                   IF NOT #found THEN
                       #VarErr := 1;                       // no feasible transfer
                   ELSIF #CurLen >= 96 THEN
                       #VarErr := 2;                       // plan longer than 96 transfers
                   ELSE
                       // ---------- apply the best (s, d) ----------
                       #si := #bS;
                       #sCol := #SrcX[#si];
                       #sRow := #SrcY[#si];
                       #sBay := #SrcB[#si];
                       #dBay := #bDb;
                       #dCol := #FreeX[#dBay, #bK];
                       #dRow := #FreeY[#dBay, #bK];
                       #eT := "Crane_MoveCost"(X0 := #cx, Y0 := #cy, B0 := #cb, X1 := #sCol, Y1 := #sRow, B1 := #sBay,
                                               MMode := #cMMode, M => #eMan);
                       #lT := "Crane_MoveCost"(X0 := #sCol, Y0 := #sRow, B0 := #sBay, X1 := #dCol, Y1 := #dRow, B1 := #dBay,
                                               MMode := #cMMode, M => #lMan);
                       #g[#dBay, #dCol, #dRow] := #g[#sBay, #sCol, #sRow];
                       #g[#sBay, #sCol, #sRow] := 0;
                       #TotT := #TotT + #eT + 200 + #lT + 200;
                       #TotM := #TotM + INT_TO_DINT(#eMan) + 1 + INT_TO_DINT(#lMan) + 1;
                       #CurLen := #CurLen + 1;
                       #CurPlan[#CurLen].Kind := #SrcKind[#si];
                       #CurPlan[#CurLen].Id := #SrcId[#si];
                       #CurPlan[#CurLen].ListIdx := #SrcIdx[#si];
                       #CurPlan[#CurLen].SrcX := INT_TO_SINT(#sCol);
                       #CurPlan[#CurLen].SrcY := INT_TO_SINT(#sRow);
                       #CurPlan[#CurLen].SrcBay := INT_TO_USINT(#sBay);
                       #CurPlan[#CurLen].DstX := INT_TO_SINT(#dCol);
                       #CurPlan[#CurLen].DstY := INT_TO_SINT(#dRow);
                       #CurPlan[#CurLen].DstBay := INT_TO_USINT(#dBay);
                       #CurPlan[#CurLen].CumT_ds := #TotT;
                       #CurPlan[#CurLen].CumM := #TotM;
                       #CurSrc[#CurLen] := #si;
                       #cx := #dCol;
                       #cy := #dRow;
                       #cb := #dBay;
                       #cG := #FreeG[#dBay, #bK];
                       #Pend[#si] := FALSE;
                       #nPend := #nPend - 1;
                   END_IF;
               END_IF;

               IF #PubPending THEN
                   // ---------- job finished: publish (World is written only here) ----------
                   #PubPending := FALSE;
                   IF #HaveBest THEN
                       FOR #i := 1 TO 96 DO
                           IF #i <= #BestLen THEN
                               "World".Plan[#i] := #BestPlan[#i];
                           ELSE
                               "World".Plan[#i] := #ZeroTr;
                           END_IF;
                       END_FOR;
                       "World".PlanLen := #BestLen;
                       "World".PlanVariant := #BestV;
                       "World".PredT_ds := #BestT;
                       "World".PredM := #BestM;
                       "World".LbT_ds := #sBaseT + #LbT;
                       "World".LbM := #sBaseM + #LbM;
                       "World".ImpEvals := #ImpEvals;
                       "World".ImpAccepts := #ImpAcc;
                       "World".SlotAccepts := #SlAcc;
                       "World".OrderFeasible := #OrderOk;
                       IF #sN > 0 THEN
                           "World".PredJ := 0.5 * (DINT_TO_REAL(#BestT) / 10.0) / (76.0 * INT_TO_REAL(#sN))
                                          + 0.5 * DINT_TO_REAL(#BestM) / (4.0 * INT_TO_REAL(#sN));
                           "World".PredJ0 := 0.5 * (DINT_TO_REAL(#GrT) / 10.0) / (76.0 * INT_TO_REAL(#sN))
                                           + 0.5 * DINT_TO_REAL(#GrM) / (4.0 * INT_TO_REAL(#sN));
                           "World".LbJ := 0.5 * (DINT_TO_REAL(#sBaseT + #LbT) / 10.0) / (76.0 * INT_TO_REAL(#sN))
                                        + 0.5 * DINT_TO_REAL(#sBaseM + #LbM) / (4.0 * INT_TO_REAL(#sN));
                       ELSE
                           "World".PredJ := 0.0;
                           "World".PredJ0 := 0.0;
                           "World".LbJ := 0.0;
                       END_IF;
                       "World".PlanValid := TRUE;
                       #Done := TRUE;
                       #ErrCode := 0;
                   ELSE
                       "World".PlanValid := FALSE;
                       "World".PlanLen := 0;
                       "World".PlanVariant := 0;
                       "World".SlotAccepts := 0;
                       "World".OrderFeasible := #OrderOk;
                       #Error := TRUE;
                       #ErrCode := #Err1;
                   END_IF;
                   #JobBusy := FALSE;
               END_IF;
           END_WHILE;
           #DiagCallMs := RUNTIME(MEM := #RtMem) * 1000.0;
           #DiagJobMs := #DiagJobMs + #DiagCallMs;
           IF #DiagCallMs > #DiagMaxCallMs THEN
               #DiagMaxCallMs := #DiagCallMs;
           END_IF;
       END_IF;
   END_REGION

   #Busy := #JobBusy;
END_FUNCTION_BLOCK

FUNCTION "CheckCmd" : Int   // FC10, SCL
TITLE = Pre-check of a crane command before OB30 issues it to FB1
{ S7_Optimized_Access := 'TRUE' }
VERSION : 0.1
// Returns 0 = OK, otherwise the alarm bit number (CONTRACT 1.4 / 3.3):
//     100 ship imbalance (alarm bit 0)      1 pick location empty
//       2 drop location occupied            9 invalid command / position
//      11 crane already carrying (lift, or MANUAL reset with a load)   12 crane is empty (put down)
//   The first failing rule decides the result.
//   Lift/put act on the CURRENT crane position (CraneX/Y/Bay); the X/Y/Bay of C are ignored.
//   Balance rule (CONTRACT 4.3 step rule): the result is OK if |L'-R'| <= BalLimit,
//   or if it is not worse than before (|L'-R'| <= |L-R|). Same for front/aft if BalMode = 1.
//   v1.5 (R2-J1): relaxed rule while "World".BalCeil > BalLimit (set by FB10 only when the ship started out
//   of balance and the list order is infeasible otherwise): while |L-R| > BalLimit, |L'-R'| <= BalCeil is OK.
   VAR_INPUT
      C : "typeCmd";   // command to check
      CraneX : SInt;   // crane position now
      CraneY : SInt;
      CraneBay : USInt;
      Carried : UInt;   // ID on the hook (0 = none)
      BalLimit : Int;   // max |L-R| (5)
      BalMode : USInt;   // 0 left/right only, 1 also front/aft
   END_VAR
   VAR_TEMP
      x : Int;
      y : Int;
      cx : Int;
      cy : Int;
      cell : UInt;
      delta : Int;   // -1 lift (container leaves the ship), +1 put
      L : Int;   // ship count x in {0,1}
      R : Int;   // ship count x in {2,3}
      F : Int;   // ship count y in 0..5
      "A" : Int;   // ship count y in 6..11
      L2 : Int;
      R2 : Int;
      F2 : Int;
      A2 : Int;
   END_VAR
BEGIN
   REGION Move and reset
       CASE #C.Cmd OF
           3:  // move to (X, Y, Bay): only the target must be a valid slot
               IF #C.X >= 0 AND #C.X <= 3 AND #C.Y >= 0 AND #C.Y <= 11 AND #C.Bay <= 1 THEN
                   #CheckCmd := 0;
               ELSE
                   #CheckCmd := 9;
               END_IF;
               RETURN;
           10: // reset of FB1: INIT may always reset (it reloads the yard and clears the hook);
               // a MANUAL reset with a container on the hook would lose it and the score counters
               IF #C.Src = 3 AND #Carried <> 0 THEN
                   #CheckCmd := 11;
               ELSE
                   #CheckCmd := 0;
               END_IF;
               RETURN;
           1, 2:
               ;   // checked below
           ELSE
               #CheckCmd := 9;
               RETURN;
       END_CASE;
   END_REGION

   REGION Lift / put: crane position and hook
       #cx := SINT_TO_INT(#CraneX);
       #cy := SINT_TO_INT(#CraneY);
       IF #cx < 0 OR #cx > 3 OR #cy < 0 OR #cy > 11 OR #CraneBay > 1 THEN
           #CheckCmd := 9;     // crane is not over a valid slot
           RETURN;
       END_IF;

       IF #CraneBay = 0 THEN
           #cell := "World".Bay0[#cx, #cy];
       ELSE
           #cell := "World".Bay1[#cx, #cy];
       END_IF;

       IF #C.Cmd = 1 THEN
           IF #Carried <> 0 THEN
               #CheckCmd := 11;    // already carrying a container
               RETURN;
           END_IF;
           IF #cell = 0 THEN
               #CheckCmd := 1;     // pick location empty
               RETURN;
           END_IF;
           #delta := -1;
       ELSE
           IF #Carried = 0 THEN
               #CheckCmd := 12;    // nothing on the hook
               RETURN;
           END_IF;
           IF #cell <> 0 THEN
               #CheckCmd := 2;     // drop location occupied
               RETURN;
           END_IF;
           #delta := 1;
       END_IF;
   END_REGION

   REGION Ship balance after the lift / put (only when it happens on the ship)
       IF #CraneBay = 0 THEN
           #L := 0; #R := 0; #F := 0; #A := 0;
           FOR #x := 0 TO 3 DO
               FOR #y := 0 TO 11 DO
                   IF "World".Bay0[#x, #y] <> 0 THEN
                       IF #x <= 1 THEN #L := #L + 1; ELSE #R := #R + 1; END_IF;
                       IF #y <= 5 THEN #F := #F + 1; ELSE #A := #A + 1; END_IF;
                   END_IF;
               END_FOR;
           END_FOR;

           #L2 := #L; #R2 := #R; #F2 := #F; #A2 := #A;
           IF #cx <= 1 THEN #L2 := #L + #delta; ELSE #R2 := #R + #delta; END_IF;
           IF #cy <= 5 THEN #F2 := #F + #delta; ELSE #A2 := #A + #delta; END_IF;

           IF ABS(#L2 - #R2) > #BalLimit AND ABS(#L2 - #R2) > ABS(#L - #R)
               AND NOT (ABS(#L - #R) > #BalLimit AND ABS(#L2 - #R2) <= "World".BalCeil)
           THEN
               #CheckCmd := 100;
               RETURN;
           END_IF;
           IF #BalMode = 1 AND ABS(#F2 - #A2) > #BalLimit AND ABS(#F2 - #A2) > ABS(#F - #A) THEN
               #CheckCmd := 100;
               RETURN;
           END_IF;
       END_IF;

       #CheckCmd := 0;
   END_REGION
END_FUNCTION

FUNCTION "Crane_MoveCost" : DInt   // FC20, SCL
TITLE = Time and manipulation cost of one crane move (CONTRACT 4.1)
{ S7_Optimized_Access := 'TRUE' }
VERSION : 0.1
// Returns the move time in DECISECONDS (DInt) from (X0,Y0,B0) to (X1,Y1,B1); output M = manipulations.
//   Global column G(x, b) = x + 6 for bay 0 (ship), x for bay 1 (yard)   (one yard bay only).
//   Same position              -> T = 0, M = 0
//   otherwise                  -> T = max(60*|dG|, 23*|dy|) ds   (6 m per column / 2.3 m per row at 1 m/s)
//   MMode 0 (spec, global X)   -> M = [dG <> 0] + [dy <> 0]
//   MMode 1 (local x)          -> M = [x1 <> x0] + [dy <> 0]
//   MMode 2 (per command, FB1) -> M = 1
//   Any other MMode is treated as 0. No range checks: callers pass valid positions
//   (the planner also uses it with synthetic columns 0..9 in bay 1 to build its cost table).
   VAR_INPUT
      X0 : Int;
      Y0 : Int;
      B0 : Int;
      X1 : Int;
      Y1 : Int;
      B1 : Int;
      MMode : Int;
   END_VAR
   VAR_OUTPUT
      "M" : Int;
   END_VAR
   VAR_TEMP
      g0 : DInt;
      g1 : DInt;
      dG : DInt;
      dY : DInt;
      tX : DInt;
      tY : DInt;
   END_VAR
BEGIN

    // Zero move: no time, no manipulation (the runtime never issues it, U6).
    IF #X0 = #X1 AND #Y0 = #Y1 AND #B0 = #B1 THEN
        #M := 0;
        #Crane_MoveCost := 0;
        RETURN;
    END_IF;

    // Global columns
    #g0 := INT_TO_DINT(#X0);
    IF #B0 = 0 THEN
        #g0 := #g0 + 6;
    END_IF;
    #g1 := INT_TO_DINT(#X1);
    IF #B1 = 0 THEN
        #g1 := #g1 + 6;
    END_IF;
    #dG := ABS(#g1 - #g0);
    #dY := ABS(INT_TO_DINT(#Y1) - INT_TO_DINT(#Y0));

    // Time: both axes travel at the same time, the longer one decides
    #tX := 60 * #dG;
    #tY := 23 * #dY;
    IF #tX >= #tY THEN
        #Crane_MoveCost := #tX;
    ELSE
        #Crane_MoveCost := #tY;
    END_IF;

    // Manipulations
    #M := 0;
    CASE #MMode OF
        1:
            IF #X1 <> #X0 THEN
                #M := #M + 1;
            END_IF;
            IF #dY <> 0 THEN
                #M := #M + 1;
            END_IF;
        2:
            #M := 1;
        ELSE
            IF #dG <> 0 THEN
                #M := #M + 1;
            END_IF;
            IF #dY <> 0 THEN
                #M := #M + 1;
            END_IF;
    END_CASE;
END_FUNCTION

FUNCTION "Crane_DropCost" : DInt   // FC21, SCL
TITLE = Weighted cost of a drop cell in the planner SLOT phase (CONTRACT 4.11)
{ S7_Optimized_Access := 'TRUE' }
VERSION : 0.1
// c(d) = W(source -> cell) + W(cell -> next source)   (second term only if HasNxt)
//   W = T [ds] + 190 * M, both from FC20 "Crane_MoveCost" (the only cost formula).
//   Python reference: tools/crane_plan.py slot_search() cost(); mirror tia-src/13_improve_mirror.py.
   VAR_INPUT
      SrcX : Int;
      SrcY : Int;
      SrcB : Int;
      CelX : Int;
      CelY : Int;
      CelB : Int;
      NxtX : Int;
      NxtY : Int;
      NxtB : Int;
      HasNxt : Bool;
      MMode : Int;
   END_VAR
   VAR_TEMP
      tA : DInt;
      mA : Int;
      wSum : DInt;
   END_VAR
BEGIN

    #tA := "Crane_MoveCost"(X0 := #SrcX, Y0 := #SrcY, B0 := #SrcB, X1 := #CelX, Y1 := #CelY, B1 := #CelB,
                            MMode := #MMode, M => #mA);
    #wSum := #tA + 190 * INT_TO_DINT(#mA);
    IF #HasNxt THEN
        #tA := "Crane_MoveCost"(X0 := #CelX, Y0 := #CelY, B0 := #CelB, X1 := #NxtX, Y1 := #NxtY, B1 := #NxtB,
                                MMode := #MMode, M => #mA);
        #wSum := #wSum + #tA + 190 * INT_TO_DINT(#mA);
    END_IF;
    #Crane_DropCost := #wSum;
END_FUNCTION

ORGANIZATION_BLOCK "Main"   // OB1, SCL, ProgramCycle
TITLE = "Main Program Sweep (Cycle)"
{ S7_Optimized_Access := 'TRUE' }
VERSION : 0.1
   VAR_INPUT
      Initial_Call : Bool;   // Initial call of this OB
      Remanence : Bool;   // =True, if remanent data are available
   END_VAR
BEGIN

    // Crane control (FB10): modes, state machine, planning, HMI interface.
    // FB1 "Crane_manipulation" is called only in OB30 "Cyclic interrupt" (1 s).
    "Crane_Control_DB"();
END_ORGANIZATION_BLOCK

ORGANIZATION_BLOCK "Cyclic interrupt"   // OB30, SCL, CyclicInterrupt
TITLE = Crane command execution (1 s cyclic interrupt)
{ S7_Optimized_Access := 'TRUE' }
VERSION : 0.1
   VAR_INPUT
      Initial_Call : Bool;   // Initial call of this OB
      Event_Count : Int;   // Events discarded
   END_VAR
   VAR_TEMP
      rc : Int;   // result of "CheckCmd"
      bitNo : Int;   // alarm bit to set in "World".Fault
      cx : Int;
      cy : Int;
      gxOld : Int;   // global column before / after a move (Bay0 x + 6, Bay1 x)
      gxNew : Int;
      cmd : "typeCmd";   // command to issue
   END_VAR
BEGIN
   // OB30 runs every 1 s (spec: "once per second"). It is the ONLY place that
   // calls FB1 "Crane_manipulation" and writes its command tags MB100..MB103.
   // FB10 "Crane_Control" (OB1) decides WHAT to do and stages it in "World".NextCmd;
   // OB30 decides WHEN: only after FB1 reported the previous command finished
   // (command_id back to 0) and only after "CheckCmd" accepted the command.
   // Order per tick (CONTRACT 3.4): 1 tick, 2 completion, 3 issue, 4 FB1 call.

   REGION 1 Tick counter and heartbeat
       "World".OB30Ticks := "World".OB30Ticks + 1;
       "HMI_IF".Heartbeat := NOT "HMI_IF".Heartbeat;
   END_REGION

   REGION 2 Has the previous command finished?
       IF "World".Busy THEN
           IF "new_command_ID" = 0 THEN
               // Spec section 3 manipulation count (shown next to FB1's MD107):
               // a move counts +1 per changed axis (x incl. bay change, y), lift / put +1, reset clears
               CASE "World".ActCmd.Cmd OF
                   1, 2:
                       "World".MSpec := "World".MSpec + 1;
                   3:
                       #gxOld := SINT_TO_INT("World".CraneX);
                       IF "World".CraneBay = 0 THEN #gxOld := #gxOld + 6; END_IF;
                       #gxNew := SINT_TO_INT("x_position");
                       IF "bay_ID" = 0 THEN #gxNew := #gxNew + 6; END_IF;
                       IF #gxNew <> #gxOld THEN "World".MSpec := "World".MSpec + 1; END_IF;
                       IF "y_position" <> "World".CraneY THEN "World".MSpec := "World".MSpec + 1; END_IF;
                   10:
                       "World".MSpec := 0;
                   ELSE
                       ;
               END_CASE;

               // FB1 finished: take over the crane position it reports
               "World".CraneX := "x_position";
               "World".CraneY := "y_position";
               "World".CraneBay := "bay_ID";

               // Effect of the command on our container model (FB1 does not track containers)
               #cx := SINT_TO_INT("World".ActCmd.X);
               #cy := SINT_TO_INT("World".ActCmd.Y);
               CASE "World".ActCmd.Cmd OF
                   1:  // lift: the container moves from the cell to the hook
                       IF #cx >= 0 AND #cx <= 3 AND #cy >= 0 AND #cy <= 11 THEN
                           IF "World".ActCmd.Bay = 0 THEN
                               "World".Carried := "World".Bay0[#cx, #cy];
                               "World".Bay0[#cx, #cy] := 0;
                           ELSIF "World".ActCmd.Bay = 1 THEN
                               "World".Carried := "World".Bay1[#cx, #cy];
                               "World".Bay1[#cx, #cy] := 0;
                           END_IF;
                       END_IF;
                   2:  // put down: the container moves from the hook to the cell
                       IF #cx >= 0 AND #cx <= 3 AND #cy >= 0 AND #cy <= 11 THEN
                           IF "World".ActCmd.Bay = 0 THEN
                               "World".Bay0[#cx, #cy] := "World".Carried;
                               "World".Carried := 0;
                           ELSIF "World".ActCmd.Bay = 1 THEN
                               "World".Bay1[#cx, #cy] := "World".Carried;
                               "World".Carried := 0;
                           END_IF;
                       END_IF;
                   3:  // move: FB1 must now report the commanded position
                       IF "World".CraneX <> "World".ActCmd.X
                           OR "World".CraneY <> "World".ActCmd.Y
                           OR "World".CraneBay <> "World".ActCmd.Bay
                       THEN
                           "World".Fault := "World".Fault OR WORD#16#4000;   // bit 14 position mismatch
                       END_IF;
                   ELSE
                       ;   // 10 reset: the crane position comes from FB1 (0,0,1)
               END_CASE;

               "World".LastDone := "World".ActCmd;
               "World".DoneSeq := "World".DoneSeq + 1;
               "World".Busy := FALSE;
               "World".BusyTicks := 0;
           ELSE
               // Still executing: watchdog
               IF "World".BusyTicks < 32000 THEN
                   "World".BusyTicks := "World".BusyTicks + 1;
               END_IF;
               IF "World".BusyTicks > "World".CfgTimeoutTicks THEN
                   "World".Fault := "World".Fault OR WORD#16#0400;           // bit 10 FB1 timeout
               END_IF;
           END_IF;
       END_IF;
   END_REGION

   REGION 3 Issue the next command (only when the previous one is done)
       // Spec 2.2: "na pocetku bloka OB30 provjeriti je li posljednja manipulacija izvrsena":
       // FB1 resets "new_command_ID" (MB103) to 0 when a command is done (checked in region 2
       // for World.Busy and here again literally, so a stray MB103 value is never overwritten).
       IF NOT "World".Busy AND "new_command_ID" = 0 AND "World".CmdReady AND "World".Permit AND "World".Fault = 0 THEN
           #cmd := "World".NextCmd;
           // Lift / put always act where the crane is now
           IF #cmd.Cmd = 1 OR #cmd.Cmd = 2 THEN
               #cmd.X := "World".CraneX;
               #cmd.Y := "World".CraneY;
               #cmd.Bay := "World".CraneBay;
           END_IF;

           // Pick not empty, drop not occupied, slot valid, ship stays balanced
           #rc := "CheckCmd"(C := #cmd,
                             CraneX := "World".CraneX,
                             CraneY := "World".CraneY,
                             CraneBay := "World".CraneBay,
                             Carried := "World".Carried,
                             BalLimit := "World".CfgBalLimit,
                             BalMode := "World".CfgBalMode);

           IF #rc = 0 THEN
               "new_x_position" := #cmd.X;
               "new_y_position" := #cmd.Y;
               "new_bay_ID" := #cmd.Bay;
               "new_command_ID" := #cmd.Cmd;
               "World".ActCmd := #cmd;
               "World".Busy := TRUE;
               "World".BusyTicks := 0;
           ELSE
               // Rejected: raise the alarm and do not issue (halts until ACK in FB10)
               IF #rc = 100 THEN
                   #bitNo := 0;
               ELSE
                   #bitNo := #rc;
               END_IF;
               IF #bitNo >= 0 AND #bitNo <= 15 THEN
                   "World".Fault := "World".Fault OR SHL(IN := WORD#16#0001, N := INT_TO_UINT(#bitNo));
               ELSE
                   "World".Fault := "World".Fault OR WORD#16#0200;           // unknown code -> bit 9
               END_IF;
               "World".FaultCmd := #cmd;
           END_IF;
           "World".CmdReady := FALSE;
       END_IF;
   END_REGION

   REGION 4 FB1 call (every tick; command 0 = nothing to do)
       "Crane_manipulation_DB"(new_x_position := "new_x_position",
                               new_y_position := "new_y_position",
                               new_bay_ID := "new_bay_ID",
                               pos_x_after_command => "x_position",
                               pos_y_after_command => "y_position",
                               bay_ID_after_command => "bay_ID",
                               number_of_manipulations => "number_of_manipulations",
                               working_time => "time",
                               command_id := "new_command_ID");
   END_REGION
END_ORGANIZATION_BLOCK

ORGANIZATION_BLOCK "Startup"   // OB100, SCL, Startup
TITLE = "Complete Restart"
{ S7_Optimized_Access := 'TRUE' }
VERSION : 0.1
   VAR_INPUT
      LostRetentive : Bool;   // True if retentive data are lost
      LostRTC : Bool;   // True if date and time are lost
   END_VAR
BEGIN
   // define the inital state of the shipyard
   "Crane_manipulation_DB".command_id := 0; // set "do nothing" command
   "Crane_manipulation_DB".current_bay_ID := 1; // the crane starting bay ID set to 1 (left of the ship)
   "Crane_manipulation_DB".current_x_position_in_bay := 0; // starting X position of the crane
   "Crane_manipulation_DB".current_y_position_in_bay := 0; // starting Y position of the crane

   //define startup command parameters
   "new_x_position" := 0; // starting X position of the crane
   "new_y_position" := 0; // starting Y position of the crane
   "new_bay_ID" := 1; // the crane starting bay ID set to 1 (left of the ship)
   "new_command_ID" := 0; // set "do nothing" command

   // reset of evaluation parameters
   "Crane_manipulation_DB".total_number_of_manipulations := 0; // reset total number of the crane manipulations
   "Crane_manipulation_DB".total_time := 0.0; // reset of total time
END_ORGANIZATION_BLOCK

(* ===== HMI "HMI_RT_1" =====
system functions are stored by id; their names below are inferred from use
connection "HMI_Connection_1": ETHERNET, S7_1500_OMS

HMI tags "Default tag table"
   "time" : Real = PLC time AT %MD112, 1 s

HMI tags "T_LinkProbe"
   "P_SwOn" : Bool = PLC HMI_IF.SwOn, 1 s

HMI tags "HMI_IF_gen"
   "SwOn" : Bool = PLC HMI_IF.SwOn AT %DB1.DBW0, 100 ms   // HMI_IF.SwOn
   "BtnInit" : Bool = PLC HMI_IF.BtnInit AT %DB1.DBW0, 100 ms   // HMI_IF.BtnInit
   "BtnAuto" : Bool = PLC HMI_IF.BtnAuto AT %DB1.DBW0, 100 ms   // HMI_IF.BtnAuto
   "BtnSemi" : Bool = PLC HMI_IF.BtnSemi AT %DB1.DBW0, 100 ms   // HMI_IF.BtnSemi
   "BtnManual" : Bool = PLC HMI_IF.BtnManual AT %DB1.DBW0, 100 ms   // HMI_IF.BtnManual
   "BtnStart" : Bool = PLC HMI_IF.BtnStart AT %DB1.DBW0, 100 ms   // HMI_IF.BtnStart
   "BtnStop" : Bool = PLC HMI_IF.BtnStop AT %DB1.DBW0, 100 ms   // HMI_IF.BtnStop
   "BtnAck" : Bool = PLC HMI_IF.BtnAck AT %DB1.DBW0, 100 ms   // HMI_IF.BtnAck
   "BtnStep" : Bool = PLC HMI_IF.BtnStep AT %DB1.DBW0, 100 ms   // HMI_IF.BtnStep
   "BtnManExec" : Bool = PLC HMI_IF.BtnManExec AT %DB1.DBW0, 100 ms   // HMI_IF.BtnManExec
   "ManCmd" : USInt = PLC HMI_IF.ManCmd AT %DB1.DBW0, 100 ms   // HMI_IF.ManCmd
   "ManX" : SInt = PLC HMI_IF.ManX AT %DB1.DBW0, 100 ms   // HMI_IF.ManX
   "ManY" : SInt = PLC HMI_IF.ManY AT %DB1.DBW0, 100 ms   // HMI_IF.ManY
   "ManBay" : USInt = PLC HMI_IF.ManBay AT %DB1.DBW0, 100 ms   // HMI_IF.ManBay
   "CfgOrderMode" : USInt = PLC HMI_IF.CfgOrderMode AT %DB1.DBW0, 100 ms   // HMI_IF.CfgOrderMode
   "CfgSemiPerTransfer" : Bool = PLC HMI_IF.CfgSemiPerTransfer AT %DB1.DBW0, 100 ms   // HMI_IF.CfgSemiPerTransfer
   "CfgBalMode" : USInt = PLC HMI_IF.CfgBalMode AT %DB1.DBW0, 100 ms   // HMI_IF.CfgBalMode
   "AlarmHmiAck" : Word = PLC HMI_IF.AlarmHmiAck AT %DB1.DBW0, 100 ms   // HMI_IF.AlarmHmiAck
   "State" : USInt = PLC HMI_IF.State AT %DB1.DBW0, 100 ms   // HMI_IF.State
   "Mode" : USInt = PLC HMI_IF.Mode AT %DB1.DBW0, 100 ms   // HMI_IF.Mode
   "LampOn" : Bool = PLC HMI_IF.LampOn AT %DB1.DBW0, 100 ms   // HMI_IF.LampOn
   "LampOff" : Bool = PLC HMI_IF.LampOff AT %DB1.DBW0, 100 ms   // HMI_IF.LampOff
   "LampReady" : Bool = PLC HMI_IF.LampReady AT %DB1.DBW0, 100 ms   // HMI_IF.LampReady
   "LampAuto" : Bool = PLC HMI_IF.LampAuto AT %DB1.DBW0, 100 ms   // HMI_IF.LampAuto
   "LampSemi" : Bool = PLC HMI_IF.LampSemi AT %DB1.DBW0, 100 ms   // HMI_IF.LampSemi
   "LampManual" : Bool = PLC HMI_IF.LampManual AT %DB1.DBW0, 100 ms   // HMI_IF.LampManual
   "LampRunning" : Bool = PLC HMI_IF.LampRunning AT %DB1.DBW0, 100 ms   // HMI_IF.LampRunning
   "LampAlarm" : Bool = PLC HMI_IF.LampAlarm AT %DB1.DBW0, 100 ms   // HMI_IF.LampAlarm
   "LampDone" : Bool = PLC HMI_IF.LampDone AT %DB1.DBW0, 100 ms   // HMI_IF.LampDone
   "Initialized" : Bool = PLC HMI_IF.Initialized AT %DB1.DBW0, 100 ms   // HMI_IF.Initialized
   "CraneBusy" : Bool = PLC HMI_IF.CraneBusy AT %DB1.DBW0, 100 ms   // HMI_IF.CraneBusy
   "Planning" : Bool = PLC HMI_IF.Planning AT %DB1.DBW0, 100 ms   // HMI_IF.Planning
   "StepWaiting" : Bool = PLC HMI_IF.StepWaiting AT %DB1.DBW0, 100 ms   // HMI_IF.StepWaiting
   "M" : UDInt = PLC HMI_IF.M AT %DB1.DBW0, 100 ms   // HMI_IF.M
   "T" : Real = PLC HMI_IF.T AT %DB1.DBW0, 100 ms   // HMI_IF.T
   "J" : Real = PLC HMI_IF.J AT %DB1.DBW0, 100 ms   // HMI_IF.J
   "MSpec" : UDInt = PLC HMI_IF.MSpec AT %DB1.DBW0, 100 ms   // HMI_IF.MSpec
   "JSpec" : Real = PLC HMI_IF.JSpec AT %DB1.DBW0, 100 ms   // HMI_IF.JSpec
   "MFb1" : UDInt = PLC HMI_IF.MFb1 AT %DB1.DBW0, 100 ms   // HMI_IF.MFb1
   "JFb1" : Real = PLC HMI_IF.JFb1 AT %DB1.DBW0, 100 ms   // HMI_IF.JFb1
   "OrderModeAct" : USInt = PLC HMI_IF.OrderModeAct AT %DB1.DBW0, 100 ms   // HMI_IF.OrderModeAct
   "OrderFallback" : Bool = PLC HMI_IF.OrderFallback AT %DB1.DBW0, 100 ms   // HMI_IF.OrderFallback
   "SlotAccepts" : DInt = PLC HMI_IF.SlotAccepts AT %DB1.DBW0, 100 ms   // HMI_IF.SlotAccepts
   "N" : Int = PLC HMI_IF.N AT %DB1.DBW0, 100 ms   // HMI_IF.N
   "PredM" : DInt = PLC HMI_IF.PredM AT %DB1.DBW0, 100 ms   // HMI_IF.PredM
   "PredT" : Real = PLC HMI_IF.PredT AT %DB1.DBW0, 100 ms   // HMI_IF.PredT
   "PredJ" : Real = PLC HMI_IF.PredJ AT %DB1.DBW0, 100 ms   // HMI_IF.PredJ
   "PredJ0" : Real = PLC HMI_IF.PredJ0 AT %DB1.DBW0, 100 ms   // HMI_IF.PredJ0
   "LbJ" : Real = PLC HMI_IF.LbJ AT %DB1.DBW0, 100 ms   // HMI_IF.LbJ
   "GapPct" : Real = PLC HMI_IF.GapPct AT %DB1.DBW0, 100 ms   // HMI_IF.GapPct
   "ImpGainPct" : Real = PLC HMI_IF.ImpGainPct AT %DB1.DBW0, 100 ms   // HMI_IF.ImpGainPct
   "ImpEvals" : DInt = PLC HMI_IF.ImpEvals AT %DB1.DBW0, 100 ms   // HMI_IF.ImpEvals
   "PlanProgress" : Int = PLC HMI_IF.PlanProgress AT %DB1.DBW0, 100 ms   // HMI_IF.PlanProgress
   "PlanVariant" : Int = PLC HMI_IF.PlanVariant AT %DB1.DBW0, 100 ms   // HMI_IF.PlanVariant
   "TrDone" : Int = PLC HMI_IF.TrDone AT %DB1.DBW0, 100 ms   // HMI_IF.TrDone
   "TrTotal" : Int = PLC HMI_IF.TrTotal AT %DB1.DBW0, 100 ms   // HMI_IF.TrTotal
   "UDone" : Int = PLC HMI_IF.UDone AT %DB1.DBW0, 100 ms   // HMI_IF.UDone
   "UTotal" : Int = PLC HMI_IF.UTotal AT %DB1.DBW0, 100 ms   // HMI_IF.UTotal
   "LDone" : Int = PLC HMI_IF.LDone AT %DB1.DBW0, 100 ms   // HMI_IF.LDone
   "LTotal" : Int = PLC HMI_IF.LTotal AT %DB1.DBW0, 100 ms   // HMI_IF.LTotal
   "CraneX" : SInt = PLC HMI_IF.CraneX AT %DB1.DBW0, 100 ms   // HMI_IF.CraneX
   "CraneY" : SInt = PLC HMI_IF.CraneY AT %DB1.DBW0, 100 ms   // HMI_IF.CraneY
   "CraneBay" : USInt = PLC HMI_IF.CraneBay AT %DB1.DBW0, 100 ms   // HMI_IF.CraneBay
   "CraneGX" : Int = PLC HMI_IF.CraneGX AT %DB1.DBW0, 100 ms   // HMI_IF.CraneGX
   "Carried" : UInt = PLC HMI_IF.Carried AT %DB1.DBW0, 100 ms   // HMI_IF.Carried
   "CurCmd" : USInt = PLC HMI_IF.CurCmd AT %DB1.DBW0, 100 ms   // HMI_IF.CurCmd
   "CurX" : SInt = PLC HMI_IF.CurX AT %DB1.DBW0, 100 ms   // HMI_IF.CurX
   "CurY" : SInt = PLC HMI_IF.CurY AT %DB1.DBW0, 100 ms   // HMI_IF.CurY
   "CurBay" : USInt = PLC HMI_IF.CurBay AT %DB1.DBW0, 100 ms   // HMI_IF.CurBay
   "CurId" : UInt = PLC HMI_IF.CurId AT %DB1.DBW0, 100 ms   // HMI_IF.CurId
   "CurKind" : USInt = PLC HMI_IF.CurKind AT %DB1.DBW0, 100 ms   // HMI_IF.CurKind
   "CurPhase" : USInt = PLC HMI_IF.CurPhase AT %DB1.DBW0, 100 ms   // HMI_IF.CurPhase
   "Cell0_00" : UInt = PLC HMI_IF.Cell0[0] AT %DB1.DBW0, 100 ms   // HMI_IF.Cell0[0]
   "Cell0_01" : UInt = PLC HMI_IF.Cell0[1] AT %DB1.DBW0, 100 ms   // HMI_IF.Cell0[1]
   "Cell0_02" : UInt = PLC HMI_IF.Cell0[2] AT %DB1.DBW0, 100 ms   // HMI_IF.Cell0[2]
   "Cell0_03" : UInt = PLC HMI_IF.Cell0[3] AT %DB1.DBW0, 100 ms   // HMI_IF.Cell0[3]
   "Cell0_04" : UInt = PLC HMI_IF.Cell0[4] AT %DB1.DBW0, 100 ms   // HMI_IF.Cell0[4]
   "Cell0_05" : UInt = PLC HMI_IF.Cell0[5] AT %DB1.DBW0, 100 ms   // HMI_IF.Cell0[5]
   "Cell0_06" : UInt = PLC HMI_IF.Cell0[6] AT %DB1.DBW0, 100 ms   // HMI_IF.Cell0[6]
   "Cell0_07" : UInt = PLC HMI_IF.Cell0[7] AT %DB1.DBW0, 100 ms   // HMI_IF.Cell0[7]
   "Cell0_08" : UInt = PLC HMI_IF.Cell0[8] AT %DB1.DBW0, 100 ms   // HMI_IF.Cell0[8]
   "Cell0_09" : UInt = PLC HMI_IF.Cell0[9] AT %DB1.DBW0, 100 ms   // HMI_IF.Cell0[9]
   "Cell0_10" : UInt = PLC HMI_IF.Cell0[10] AT %DB1.DBW0, 100 ms   // HMI_IF.Cell0[10]
   "Cell0_11" : UInt = PLC HMI_IF.Cell0[11] AT %DB1.DBW0, 100 ms   // HMI_IF.Cell0[11]
   "Cell0_12" : UInt = PLC HMI_IF.Cell0[12] AT %DB1.DBW0, 100 ms   // HMI_IF.Cell0[12]
   "Cell0_13" : UInt = PLC HMI_IF.Cell0[13] AT %DB1.DBW0, 100 ms   // HMI_IF.Cell0[13]
   "Cell0_14" : UInt = PLC HMI_IF.Cell0[14] AT %DB1.DBW0, 100 ms   // HMI_IF.Cell0[14]
   "Cell0_15" : UInt = PLC HMI_IF.Cell0[15] AT %DB1.DBW0, 100 ms   // HMI_IF.Cell0[15]
   "Cell0_16" : UInt = PLC HMI_IF.Cell0[16] AT %DB1.DBW0, 100 ms   // HMI_IF.Cell0[16]
   "Cell0_17" : UInt = PLC HMI_IF.Cell0[17] AT %DB1.DBW0, 100 ms   // HMI_IF.Cell0[17]
   "Cell0_18" : UInt = PLC HMI_IF.Cell0[18] AT %DB1.DBW0, 100 ms   // HMI_IF.Cell0[18]
   "Cell0_19" : UInt = PLC HMI_IF.Cell0[19] AT %DB1.DBW0, 100 ms   // HMI_IF.Cell0[19]
   "Cell0_20" : UInt = PLC HMI_IF.Cell0[20] AT %DB1.DBW0, 100 ms   // HMI_IF.Cell0[20]
   "Cell0_21" : UInt = PLC HMI_IF.Cell0[21] AT %DB1.DBW0, 100 ms   // HMI_IF.Cell0[21]
   "Cell0_22" : UInt = PLC HMI_IF.Cell0[22] AT %DB1.DBW0, 100 ms   // HMI_IF.Cell0[22]
   "Cell0_23" : UInt = PLC HMI_IF.Cell0[23] AT %DB1.DBW0, 100 ms   // HMI_IF.Cell0[23]
   "Cell0_24" : UInt = PLC HMI_IF.Cell0[24] AT %DB1.DBW0, 100 ms   // HMI_IF.Cell0[24]
   "Cell0_25" : UInt = PLC HMI_IF.Cell0[25] AT %DB1.DBW0, 100 ms   // HMI_IF.Cell0[25]
   "Cell0_26" : UInt = PLC HMI_IF.Cell0[26] AT %DB1.DBW0, 100 ms   // HMI_IF.Cell0[26]
   "Cell0_27" : UInt = PLC HMI_IF.Cell0[27] AT %DB1.DBW0, 100 ms   // HMI_IF.Cell0[27]
   "Cell0_28" : UInt = PLC HMI_IF.Cell0[28] AT %DB1.DBW0, 100 ms   // HMI_IF.Cell0[28]
   "Cell0_29" : UInt = PLC HMI_IF.Cell0[29] AT %DB1.DBW0, 100 ms   // HMI_IF.Cell0[29]
   "Cell0_30" : UInt = PLC HMI_IF.Cell0[30] AT %DB1.DBW0, 100 ms   // HMI_IF.Cell0[30]
   "Cell0_31" : UInt = PLC HMI_IF.Cell0[31] AT %DB1.DBW0, 100 ms   // HMI_IF.Cell0[31]
   "Cell0_32" : UInt = PLC HMI_IF.Cell0[32] AT %DB1.DBW0, 100 ms   // HMI_IF.Cell0[32]
   "Cell0_33" : UInt = PLC HMI_IF.Cell0[33] AT %DB1.DBW0, 100 ms   // HMI_IF.Cell0[33]
   "Cell0_34" : UInt = PLC HMI_IF.Cell0[34] AT %DB1.DBW0, 100 ms   // HMI_IF.Cell0[34]
   "Cell0_35" : UInt = PLC HMI_IF.Cell0[35] AT %DB1.DBW0, 100 ms   // HMI_IF.Cell0[35]
   "Cell0_36" : UInt = PLC HMI_IF.Cell0[36] AT %DB1.DBW0, 100 ms   // HMI_IF.Cell0[36]
   "Cell0_37" : UInt = PLC HMI_IF.Cell0[37] AT %DB1.DBW0, 100 ms   // HMI_IF.Cell0[37]
   "Cell0_38" : UInt = PLC HMI_IF.Cell0[38] AT %DB1.DBW0, 100 ms   // HMI_IF.Cell0[38]
   "Cell0_39" : UInt = PLC HMI_IF.Cell0[39] AT %DB1.DBW0, 100 ms   // HMI_IF.Cell0[39]
   "Cell0_40" : UInt = PLC HMI_IF.Cell0[40] AT %DB1.DBW0, 100 ms   // HMI_IF.Cell0[40]
   "Cell0_41" : UInt = PLC HMI_IF.Cell0[41] AT %DB1.DBW0, 100 ms   // HMI_IF.Cell0[41]
   "Cell0_42" : UInt = PLC HMI_IF.Cell0[42] AT %DB1.DBW0, 100 ms   // HMI_IF.Cell0[42]
   "Cell0_43" : UInt = PLC HMI_IF.Cell0[43] AT %DB1.DBW0, 100 ms   // HMI_IF.Cell0[43]
   "Cell0_44" : UInt = PLC HMI_IF.Cell0[44] AT %DB1.DBW0, 100 ms   // HMI_IF.Cell0[44]
   "Cell0_45" : UInt = PLC HMI_IF.Cell0[45] AT %DB1.DBW0, 100 ms   // HMI_IF.Cell0[45]
   "Cell0_46" : UInt = PLC HMI_IF.Cell0[46] AT %DB1.DBW0, 100 ms   // HMI_IF.Cell0[46]
   "Cell0_47" : UInt = PLC HMI_IF.Cell0[47] AT %DB1.DBW0, 100 ms   // HMI_IF.Cell0[47]
   "Cell1_00" : UInt = PLC HMI_IF.Cell1[0] AT %DB1.DBW0, 100 ms   // HMI_IF.Cell1[0]
   "Cell1_01" : UInt = PLC HMI_IF.Cell1[1] AT %DB1.DBW0, 100 ms   // HMI_IF.Cell1[1]
   "Cell1_02" : UInt = PLC HMI_IF.Cell1[2] AT %DB1.DBW0, 100 ms   // HMI_IF.Cell1[2]
   "Cell1_03" : UInt = PLC HMI_IF.Cell1[3] AT %DB1.DBW0, 100 ms   // HMI_IF.Cell1[3]
   "Cell1_04" : UInt = PLC HMI_IF.Cell1[4] AT %DB1.DBW0, 100 ms   // HMI_IF.Cell1[4]
   "Cell1_05" : UInt = PLC HMI_IF.Cell1[5] AT %DB1.DBW0, 100 ms   // HMI_IF.Cell1[5]
   "Cell1_06" : UInt = PLC HMI_IF.Cell1[6] AT %DB1.DBW0, 100 ms   // HMI_IF.Cell1[6]
   "Cell1_07" : UInt = PLC HMI_IF.Cell1[7] AT %DB1.DBW0, 100 ms   // HMI_IF.Cell1[7]
   "Cell1_08" : UInt = PLC HMI_IF.Cell1[8] AT %DB1.DBW0, 100 ms   // HMI_IF.Cell1[8]
   "Cell1_09" : UInt = PLC HMI_IF.Cell1[9] AT %DB1.DBW0, 100 ms   // HMI_IF.Cell1[9]
   "Cell1_10" : UInt = PLC HMI_IF.Cell1[10] AT %DB1.DBW0, 100 ms   // HMI_IF.Cell1[10]
   "Cell1_11" : UInt = PLC HMI_IF.Cell1[11] AT %DB1.DBW0, 100 ms   // HMI_IF.Cell1[11]
   "Cell1_12" : UInt = PLC HMI_IF.Cell1[12] AT %DB1.DBW0, 100 ms   // HMI_IF.Cell1[12]
   "Cell1_13" : UInt = PLC HMI_IF.Cell1[13] AT %DB1.DBW0, 100 ms   // HMI_IF.Cell1[13]
   "Cell1_14" : UInt = PLC HMI_IF.Cell1[14] AT %DB1.DBW0, 100 ms   // HMI_IF.Cell1[14]
   "Cell1_15" : UInt = PLC HMI_IF.Cell1[15] AT %DB1.DBW0, 100 ms   // HMI_IF.Cell1[15]
   "Cell1_16" : UInt = PLC HMI_IF.Cell1[16] AT %DB1.DBW0, 100 ms   // HMI_IF.Cell1[16]
   "Cell1_17" : UInt = PLC HMI_IF.Cell1[17] AT %DB1.DBW0, 100 ms   // HMI_IF.Cell1[17]
   "Cell1_18" : UInt = PLC HMI_IF.Cell1[18] AT %DB1.DBW0, 100 ms   // HMI_IF.Cell1[18]
   "Cell1_19" : UInt = PLC HMI_IF.Cell1[19] AT %DB1.DBW0, 100 ms   // HMI_IF.Cell1[19]
   "Cell1_20" : UInt = PLC HMI_IF.Cell1[20] AT %DB1.DBW0, 100 ms   // HMI_IF.Cell1[20]
   "Cell1_21" : UInt = PLC HMI_IF.Cell1[21] AT %DB1.DBW0, 100 ms   // HMI_IF.Cell1[21]
   "Cell1_22" : UInt = PLC HMI_IF.Cell1[22] AT %DB1.DBW0, 100 ms   // HMI_IF.Cell1[22]
   "Cell1_23" : UInt = PLC HMI_IF.Cell1[23] AT %DB1.DBW0, 100 ms   // HMI_IF.Cell1[23]
   "Cell1_24" : UInt = PLC HMI_IF.Cell1[24] AT %DB1.DBW0, 100 ms   // HMI_IF.Cell1[24]
   "Cell1_25" : UInt = PLC HMI_IF.Cell1[25] AT %DB1.DBW0, 100 ms   // HMI_IF.Cell1[25]
   "Cell1_26" : UInt = PLC HMI_IF.Cell1[26] AT %DB1.DBW0, 100 ms   // HMI_IF.Cell1[26]
   "Cell1_27" : UInt = PLC HMI_IF.Cell1[27] AT %DB1.DBW0, 100 ms   // HMI_IF.Cell1[27]
   "Cell1_28" : UInt = PLC HMI_IF.Cell1[28] AT %DB1.DBW0, 100 ms   // HMI_IF.Cell1[28]
   "Cell1_29" : UInt = PLC HMI_IF.Cell1[29] AT %DB1.DBW0, 100 ms   // HMI_IF.Cell1[29]
   "Cell1_30" : UInt = PLC HMI_IF.Cell1[30] AT %DB1.DBW0, 100 ms   // HMI_IF.Cell1[30]
   "Cell1_31" : UInt = PLC HMI_IF.Cell1[31] AT %DB1.DBW0, 100 ms   // HMI_IF.Cell1[31]
   "Cell1_32" : UInt = PLC HMI_IF.Cell1[32] AT %DB1.DBW0, 100 ms   // HMI_IF.Cell1[32]
   "Cell1_33" : UInt = PLC HMI_IF.Cell1[33] AT %DB1.DBW0, 100 ms   // HMI_IF.Cell1[33]
   "Cell1_34" : UInt = PLC HMI_IF.Cell1[34] AT %DB1.DBW0, 100 ms   // HMI_IF.Cell1[34]
   "Cell1_35" : UInt = PLC HMI_IF.Cell1[35] AT %DB1.DBW0, 100 ms   // HMI_IF.Cell1[35]
   "Cell1_36" : UInt = PLC HMI_IF.Cell1[36] AT %DB1.DBW0, 100 ms   // HMI_IF.Cell1[36]
   "Cell1_37" : UInt = PLC HMI_IF.Cell1[37] AT %DB1.DBW0, 100 ms   // HMI_IF.Cell1[37]
   "Cell1_38" : UInt = PLC HMI_IF.Cell1[38] AT %DB1.DBW0, 100 ms   // HMI_IF.Cell1[38]
   "Cell1_39" : UInt = PLC HMI_IF.Cell1[39] AT %DB1.DBW0, 100 ms   // HMI_IF.Cell1[39]
   "Cell1_40" : UInt = PLC HMI_IF.Cell1[40] AT %DB1.DBW0, 100 ms   // HMI_IF.Cell1[40]
   "Cell1_41" : UInt = PLC HMI_IF.Cell1[41] AT %DB1.DBW0, 100 ms   // HMI_IF.Cell1[41]
   "Cell1_42" : UInt = PLC HMI_IF.Cell1[42] AT %DB1.DBW0, 100 ms   // HMI_IF.Cell1[42]
   "Cell1_43" : UInt = PLC HMI_IF.Cell1[43] AT %DB1.DBW0, 100 ms   // HMI_IF.Cell1[43]
   "Cell1_44" : UInt = PLC HMI_IF.Cell1[44] AT %DB1.DBW0, 100 ms   // HMI_IF.Cell1[44]
   "Cell1_45" : UInt = PLC HMI_IF.Cell1[45] AT %DB1.DBW0, 100 ms   // HMI_IF.Cell1[45]
   "Cell1_46" : UInt = PLC HMI_IF.Cell1[46] AT %DB1.DBW0, 100 ms   // HMI_IF.Cell1[46]
   "Cell1_47" : UInt = PLC HMI_IF.Cell1[47] AT %DB1.DBW0, 100 ms   // HMI_IF.Cell1[47]
   "CellSt0_00" : USInt = PLC HMI_IF.CellSt0[0] AT %DB1.DBW0, 100 ms   // HMI_IF.CellSt0[0]
   "CellSt0_01" : USInt = PLC HMI_IF.CellSt0[1] AT %DB1.DBW0, 100 ms   // HMI_IF.CellSt0[1]
   "CellSt0_02" : USInt = PLC HMI_IF.CellSt0[2] AT %DB1.DBW0, 100 ms   // HMI_IF.CellSt0[2]
   "CellSt0_03" : USInt = PLC HMI_IF.CellSt0[3] AT %DB1.DBW0, 100 ms   // HMI_IF.CellSt0[3]
   "CellSt0_04" : USInt = PLC HMI_IF.CellSt0[4] AT %DB1.DBW0, 100 ms   // HMI_IF.CellSt0[4]
   "CellSt0_05" : USInt = PLC HMI_IF.CellSt0[5] AT %DB1.DBW0, 100 ms   // HMI_IF.CellSt0[5]
   "CellSt0_06" : USInt = PLC HMI_IF.CellSt0[6] AT %DB1.DBW0, 100 ms   // HMI_IF.CellSt0[6]
   "CellSt0_07" : USInt = PLC HMI_IF.CellSt0[7] AT %DB1.DBW0, 100 ms   // HMI_IF.CellSt0[7]
   "CellSt0_08" : USInt = PLC HMI_IF.CellSt0[8] AT %DB1.DBW0, 100 ms   // HMI_IF.CellSt0[8]
   "CellSt0_09" : USInt = PLC HMI_IF.CellSt0[9] AT %DB1.DBW0, 100 ms   // HMI_IF.CellSt0[9]
   "CellSt0_10" : USInt = PLC HMI_IF.CellSt0[10] AT %DB1.DBW0, 100 ms   // HMI_IF.CellSt0[10]
   "CellSt0_11" : USInt = PLC HMI_IF.CellSt0[11] AT %DB1.DBW0, 100 ms   // HMI_IF.CellSt0[11]
   "CellSt0_12" : USInt = PLC HMI_IF.CellSt0[12] AT %DB1.DBW0, 100 ms   // HMI_IF.CellSt0[12]
   "CellSt0_13" : USInt = PLC HMI_IF.CellSt0[13] AT %DB1.DBW0, 100 ms   // HMI_IF.CellSt0[13]
   "CellSt0_14" : USInt = PLC HMI_IF.CellSt0[14] AT %DB1.DBW0, 100 ms   // HMI_IF.CellSt0[14]
   "CellSt0_15" : USInt = PLC HMI_IF.CellSt0[15] AT %DB1.DBW0, 100 ms   // HMI_IF.CellSt0[15]
   "CellSt0_16" : USInt = PLC HMI_IF.CellSt0[16] AT %DB1.DBW0, 100 ms   // HMI_IF.CellSt0[16]
   "CellSt0_17" : USInt = PLC HMI_IF.CellSt0[17] AT %DB1.DBW0, 100 ms   // HMI_IF.CellSt0[17]
   "CellSt0_18" : USInt = PLC HMI_IF.CellSt0[18] AT %DB1.DBW0, 100 ms   // HMI_IF.CellSt0[18]
   "CellSt0_19" : USInt = PLC HMI_IF.CellSt0[19] AT %DB1.DBW0, 100 ms   // HMI_IF.CellSt0[19]
   "CellSt0_20" : USInt = PLC HMI_IF.CellSt0[20] AT %DB1.DBW0, 100 ms   // HMI_IF.CellSt0[20]
   "CellSt0_21" : USInt = PLC HMI_IF.CellSt0[21] AT %DB1.DBW0, 100 ms   // HMI_IF.CellSt0[21]
   "CellSt0_22" : USInt = PLC HMI_IF.CellSt0[22] AT %DB1.DBW0, 100 ms   // HMI_IF.CellSt0[22]
   "CellSt0_23" : USInt = PLC HMI_IF.CellSt0[23] AT %DB1.DBW0, 100 ms   // HMI_IF.CellSt0[23]
   "CellSt0_24" : USInt = PLC HMI_IF.CellSt0[24] AT %DB1.DBW0, 100 ms   // HMI_IF.CellSt0[24]
   "CellSt0_25" : USInt = PLC HMI_IF.CellSt0[25] AT %DB1.DBW0, 100 ms   // HMI_IF.CellSt0[25]
   "CellSt0_26" : USInt = PLC HMI_IF.CellSt0[26] AT %DB1.DBW0, 100 ms   // HMI_IF.CellSt0[26]
   "CellSt0_27" : USInt = PLC HMI_IF.CellSt0[27] AT %DB1.DBW0, 100 ms   // HMI_IF.CellSt0[27]
   "CellSt0_28" : USInt = PLC HMI_IF.CellSt0[28] AT %DB1.DBW0, 100 ms   // HMI_IF.CellSt0[28]
   "CellSt0_29" : USInt = PLC HMI_IF.CellSt0[29] AT %DB1.DBW0, 100 ms   // HMI_IF.CellSt0[29]
   "CellSt0_30" : USInt = PLC HMI_IF.CellSt0[30] AT %DB1.DBW0, 100 ms   // HMI_IF.CellSt0[30]
   "CellSt0_31" : USInt = PLC HMI_IF.CellSt0[31] AT %DB1.DBW0, 100 ms   // HMI_IF.CellSt0[31]
   "CellSt0_32" : USInt = PLC HMI_IF.CellSt0[32] AT %DB1.DBW0, 100 ms   // HMI_IF.CellSt0[32]
   "CellSt0_33" : USInt = PLC HMI_IF.CellSt0[33] AT %DB1.DBW0, 100 ms   // HMI_IF.CellSt0[33]
   "CellSt0_34" : USInt = PLC HMI_IF.CellSt0[34] AT %DB1.DBW0, 100 ms   // HMI_IF.CellSt0[34]
   "CellSt0_35" : USInt = PLC HMI_IF.CellSt0[35] AT %DB1.DBW0, 100 ms   // HMI_IF.CellSt0[35]
   "CellSt0_36" : USInt = PLC HMI_IF.CellSt0[36] AT %DB1.DBW0, 100 ms   // HMI_IF.CellSt0[36]
   "CellSt0_37" : USInt = PLC HMI_IF.CellSt0[37] AT %DB1.DBW0, 100 ms   // HMI_IF.CellSt0[37]
   "CellSt0_38" : USInt = PLC HMI_IF.CellSt0[38] AT %DB1.DBW0, 100 ms   // HMI_IF.CellSt0[38]
   "CellSt0_39" : USInt = PLC HMI_IF.CellSt0[39] AT %DB1.DBW0, 100 ms   // HMI_IF.CellSt0[39]
   "CellSt0_40" : USInt = PLC HMI_IF.CellSt0[40] AT %DB1.DBW0, 100 ms   // HMI_IF.CellSt0[40]
   "CellSt0_41" : USInt = PLC HMI_IF.CellSt0[41] AT %DB1.DBW0, 100 ms   // HMI_IF.CellSt0[41]
   "CellSt0_42" : USInt = PLC HMI_IF.CellSt0[42] AT %DB1.DBW0, 100 ms   // HMI_IF.CellSt0[42]
   "CellSt0_43" : USInt = PLC HMI_IF.CellSt0[43] AT %DB1.DBW0, 100 ms   // HMI_IF.CellSt0[43]
   "CellSt0_44" : USInt = PLC HMI_IF.CellSt0[44] AT %DB1.DBW0, 100 ms   // HMI_IF.CellSt0[44]
   "CellSt0_45" : USInt = PLC HMI_IF.CellSt0[45] AT %DB1.DBW0, 100 ms   // HMI_IF.CellSt0[45]
   "CellSt0_46" : USInt = PLC HMI_IF.CellSt0[46] AT %DB1.DBW0, 100 ms   // HMI_IF.CellSt0[46]
   "CellSt0_47" : USInt = PLC HMI_IF.CellSt0[47] AT %DB1.DBW0, 100 ms   // HMI_IF.CellSt0[47]
   "CellSt1_00" : USInt = PLC HMI_IF.CellSt1[0] AT %DB1.DBW0, 100 ms   // HMI_IF.CellSt1[0]
   "CellSt1_01" : USInt = PLC HMI_IF.CellSt1[1] AT %DB1.DBW0, 100 ms   // HMI_IF.CellSt1[1]
   "CellSt1_02" : USInt = PLC HMI_IF.CellSt1[2] AT %DB1.DBW0, 100 ms   // HMI_IF.CellSt1[2]
   "CellSt1_03" : USInt = PLC HMI_IF.CellSt1[3] AT %DB1.DBW0, 100 ms   // HMI_IF.CellSt1[3]
   "CellSt1_04" : USInt = PLC HMI_IF.CellSt1[4] AT %DB1.DBW0, 100 ms   // HMI_IF.CellSt1[4]
   "CellSt1_05" : USInt = PLC HMI_IF.CellSt1[5] AT %DB1.DBW0, 100 ms   // HMI_IF.CellSt1[5]
   "CellSt1_06" : USInt = PLC HMI_IF.CellSt1[6] AT %DB1.DBW0, 100 ms   // HMI_IF.CellSt1[6]
   "CellSt1_07" : USInt = PLC HMI_IF.CellSt1[7] AT %DB1.DBW0, 100 ms   // HMI_IF.CellSt1[7]
   "CellSt1_08" : USInt = PLC HMI_IF.CellSt1[8] AT %DB1.DBW0, 100 ms   // HMI_IF.CellSt1[8]
   "CellSt1_09" : USInt = PLC HMI_IF.CellSt1[9] AT %DB1.DBW0, 100 ms   // HMI_IF.CellSt1[9]
   "CellSt1_10" : USInt = PLC HMI_IF.CellSt1[10] AT %DB1.DBW0, 100 ms   // HMI_IF.CellSt1[10]
   "CellSt1_11" : USInt = PLC HMI_IF.CellSt1[11] AT %DB1.DBW0, 100 ms   // HMI_IF.CellSt1[11]
   "CellSt1_12" : USInt = PLC HMI_IF.CellSt1[12] AT %DB1.DBW0, 100 ms   // HMI_IF.CellSt1[12]
   "CellSt1_13" : USInt = PLC HMI_IF.CellSt1[13] AT %DB1.DBW0, 100 ms   // HMI_IF.CellSt1[13]
   "CellSt1_14" : USInt = PLC HMI_IF.CellSt1[14] AT %DB1.DBW0, 100 ms   // HMI_IF.CellSt1[14]
   "CellSt1_15" : USInt = PLC HMI_IF.CellSt1[15] AT %DB1.DBW0, 100 ms   // HMI_IF.CellSt1[15]
   "CellSt1_16" : USInt = PLC HMI_IF.CellSt1[16] AT %DB1.DBW0, 100 ms   // HMI_IF.CellSt1[16]
   "CellSt1_17" : USInt = PLC HMI_IF.CellSt1[17] AT %DB1.DBW0, 100 ms   // HMI_IF.CellSt1[17]
   "CellSt1_18" : USInt = PLC HMI_IF.CellSt1[18] AT %DB1.DBW0, 100 ms   // HMI_IF.CellSt1[18]
   "CellSt1_19" : USInt = PLC HMI_IF.CellSt1[19] AT %DB1.DBW0, 100 ms   // HMI_IF.CellSt1[19]
   "CellSt1_20" : USInt = PLC HMI_IF.CellSt1[20] AT %DB1.DBW0, 100 ms   // HMI_IF.CellSt1[20]
   "CellSt1_21" : USInt = PLC HMI_IF.CellSt1[21] AT %DB1.DBW0, 100 ms   // HMI_IF.CellSt1[21]
   "CellSt1_22" : USInt = PLC HMI_IF.CellSt1[22] AT %DB1.DBW0, 100 ms   // HMI_IF.CellSt1[22]
   "CellSt1_23" : USInt = PLC HMI_IF.CellSt1[23] AT %DB1.DBW0, 100 ms   // HMI_IF.CellSt1[23]
   "CellSt1_24" : USInt = PLC HMI_IF.CellSt1[24] AT %DB1.DBW0, 100 ms   // HMI_IF.CellSt1[24]
   "CellSt1_25" : USInt = PLC HMI_IF.CellSt1[25] AT %DB1.DBW0, 100 ms   // HMI_IF.CellSt1[25]
   "CellSt1_26" : USInt = PLC HMI_IF.CellSt1[26] AT %DB1.DBW0, 100 ms   // HMI_IF.CellSt1[26]
   "CellSt1_27" : USInt = PLC HMI_IF.CellSt1[27] AT %DB1.DBW0, 100 ms   // HMI_IF.CellSt1[27]
   "CellSt1_28" : USInt = PLC HMI_IF.CellSt1[28] AT %DB1.DBW0, 100 ms   // HMI_IF.CellSt1[28]
   "CellSt1_29" : USInt = PLC HMI_IF.CellSt1[29] AT %DB1.DBW0, 100 ms   // HMI_IF.CellSt1[29]
   "CellSt1_30" : USInt = PLC HMI_IF.CellSt1[30] AT %DB1.DBW0, 100 ms   // HMI_IF.CellSt1[30]
   "CellSt1_31" : USInt = PLC HMI_IF.CellSt1[31] AT %DB1.DBW0, 100 ms   // HMI_IF.CellSt1[31]
   "CellSt1_32" : USInt = PLC HMI_IF.CellSt1[32] AT %DB1.DBW0, 100 ms   // HMI_IF.CellSt1[32]
   "CellSt1_33" : USInt = PLC HMI_IF.CellSt1[33] AT %DB1.DBW0, 100 ms   // HMI_IF.CellSt1[33]
   "CellSt1_34" : USInt = PLC HMI_IF.CellSt1[34] AT %DB1.DBW0, 100 ms   // HMI_IF.CellSt1[34]
   "CellSt1_35" : USInt = PLC HMI_IF.CellSt1[35] AT %DB1.DBW0, 100 ms   // HMI_IF.CellSt1[35]
   "CellSt1_36" : USInt = PLC HMI_IF.CellSt1[36] AT %DB1.DBW0, 100 ms   // HMI_IF.CellSt1[36]
   "CellSt1_37" : USInt = PLC HMI_IF.CellSt1[37] AT %DB1.DBW0, 100 ms   // HMI_IF.CellSt1[37]
   "CellSt1_38" : USInt = PLC HMI_IF.CellSt1[38] AT %DB1.DBW0, 100 ms   // HMI_IF.CellSt1[38]
   "CellSt1_39" : USInt = PLC HMI_IF.CellSt1[39] AT %DB1.DBW0, 100 ms   // HMI_IF.CellSt1[39]
   "CellSt1_40" : USInt = PLC HMI_IF.CellSt1[40] AT %DB1.DBW0, 100 ms   // HMI_IF.CellSt1[40]
   "CellSt1_41" : USInt = PLC HMI_IF.CellSt1[41] AT %DB1.DBW0, 100 ms   // HMI_IF.CellSt1[41]
   "CellSt1_42" : USInt = PLC HMI_IF.CellSt1[42] AT %DB1.DBW0, 100 ms   // HMI_IF.CellSt1[42]
   "CellSt1_43" : USInt = PLC HMI_IF.CellSt1[43] AT %DB1.DBW0, 100 ms   // HMI_IF.CellSt1[43]
   "CellSt1_44" : USInt = PLC HMI_IF.CellSt1[44] AT %DB1.DBW0, 100 ms   // HMI_IF.CellSt1[44]
   "CellSt1_45" : USInt = PLC HMI_IF.CellSt1[45] AT %DB1.DBW0, 100 ms   // HMI_IF.CellSt1[45]
   "CellSt1_46" : USInt = PLC HMI_IF.CellSt1[46] AT %DB1.DBW0, 100 ms   // HMI_IF.CellSt1[46]
   "CellSt1_47" : USInt = PLC HMI_IF.CellSt1[47] AT %DB1.DBW0, 100 ms   // HMI_IF.CellSt1[47]
   "UList_01" : UInt = PLC HMI_IF.UList[1] AT %DB1.DBW0, 100 ms   // HMI_IF.UList[1]
   "UList_02" : UInt = PLC HMI_IF.UList[2] AT %DB1.DBW0, 100 ms   // HMI_IF.UList[2]
   "UList_03" : UInt = PLC HMI_IF.UList[3] AT %DB1.DBW0, 100 ms   // HMI_IF.UList[3]
   "UList_04" : UInt = PLC HMI_IF.UList[4] AT %DB1.DBW0, 100 ms   // HMI_IF.UList[4]
   "UList_05" : UInt = PLC HMI_IF.UList[5] AT %DB1.DBW0, 100 ms   // HMI_IF.UList[5]
   "UList_06" : UInt = PLC HMI_IF.UList[6] AT %DB1.DBW0, 100 ms   // HMI_IF.UList[6]
   "UList_07" : UInt = PLC HMI_IF.UList[7] AT %DB1.DBW0, 100 ms   // HMI_IF.UList[7]
   "UList_08" : UInt = PLC HMI_IF.UList[8] AT %DB1.DBW0, 100 ms   // HMI_IF.UList[8]
   "UList_09" : UInt = PLC HMI_IF.UList[9] AT %DB1.DBW0, 100 ms   // HMI_IF.UList[9]
   "UList_10" : UInt = PLC HMI_IF.UList[10] AT %DB1.DBW0, 100 ms   // HMI_IF.UList[10]
   "UList_11" : UInt = PLC HMI_IF.UList[11] AT %DB1.DBW0, 100 ms   // HMI_IF.UList[11]
   "UList_12" : UInt = PLC HMI_IF.UList[12] AT %DB1.DBW0, 100 ms   // HMI_IF.UList[12]
   "UList_13" : UInt = PLC HMI_IF.UList[13] AT %DB1.DBW0, 100 ms   // HMI_IF.UList[13]
   "UList_14" : UInt = PLC HMI_IF.UList[14] AT %DB1.DBW0, 100 ms   // HMI_IF.UList[14]
   "UList_15" : UInt = PLC HMI_IF.UList[15] AT %DB1.DBW0, 100 ms   // HMI_IF.UList[15]
   "UList_16" : UInt = PLC HMI_IF.UList[16] AT %DB1.DBW0, 100 ms   // HMI_IF.UList[16]
   "UList_17" : UInt = PLC HMI_IF.UList[17] AT %DB1.DBW0, 100 ms   // HMI_IF.UList[17]
   "UList_18" : UInt = PLC HMI_IF.UList[18] AT %DB1.DBW0, 100 ms   // HMI_IF.UList[18]
   "UList_19" : UInt = PLC HMI_IF.UList[19] AT %DB1.DBW0, 100 ms   // HMI_IF.UList[19]
   "UList_20" : UInt = PLC HMI_IF.UList[20] AT %DB1.DBW0, 100 ms   // HMI_IF.UList[20]
   "UList_21" : UInt = PLC HMI_IF.UList[21] AT %DB1.DBW0, 100 ms   // HMI_IF.UList[21]
   "UList_22" : UInt = PLC HMI_IF.UList[22] AT %DB1.DBW0, 100 ms   // HMI_IF.UList[22]
   "UList_23" : UInt = PLC HMI_IF.UList[23] AT %DB1.DBW0, 100 ms   // HMI_IF.UList[23]
   "UList_24" : UInt = PLC HMI_IF.UList[24] AT %DB1.DBW0, 100 ms   // HMI_IF.UList[24]
   "UList_25" : UInt = PLC HMI_IF.UList[25] AT %DB1.DBW0, 100 ms   // HMI_IF.UList[25]
   "UList_26" : UInt = PLC HMI_IF.UList[26] AT %DB1.DBW0, 100 ms   // HMI_IF.UList[26]
   "UList_27" : UInt = PLC HMI_IF.UList[27] AT %DB1.DBW0, 100 ms   // HMI_IF.UList[27]
   "UList_28" : UInt = PLC HMI_IF.UList[28] AT %DB1.DBW0, 100 ms   // HMI_IF.UList[28]
   "UList_29" : UInt = PLC HMI_IF.UList[29] AT %DB1.DBW0, 100 ms   // HMI_IF.UList[29]
   "UList_30" : UInt = PLC HMI_IF.UList[30] AT %DB1.DBW0, 100 ms   // HMI_IF.UList[30]
   "UList_31" : UInt = PLC HMI_IF.UList[31] AT %DB1.DBW0, 100 ms   // HMI_IF.UList[31]
   "UList_32" : UInt = PLC HMI_IF.UList[32] AT %DB1.DBW0, 100 ms   // HMI_IF.UList[32]
   "UList_33" : UInt = PLC HMI_IF.UList[33] AT %DB1.DBW0, 100 ms   // HMI_IF.UList[33]
   "UList_34" : UInt = PLC HMI_IF.UList[34] AT %DB1.DBW0, 100 ms   // HMI_IF.UList[34]
   "UList_35" : UInt = PLC HMI_IF.UList[35] AT %DB1.DBW0, 100 ms   // HMI_IF.UList[35]
   "UList_36" : UInt = PLC HMI_IF.UList[36] AT %DB1.DBW0, 100 ms   // HMI_IF.UList[36]
   "UList_37" : UInt = PLC HMI_IF.UList[37] AT %DB1.DBW0, 100 ms   // HMI_IF.UList[37]
   "UList_38" : UInt = PLC HMI_IF.UList[38] AT %DB1.DBW0, 100 ms   // HMI_IF.UList[38]
   "UList_39" : UInt = PLC HMI_IF.UList[39] AT %DB1.DBW0, 100 ms   // HMI_IF.UList[39]
   "UList_40" : UInt = PLC HMI_IF.UList[40] AT %DB1.DBW0, 100 ms   // HMI_IF.UList[40]
   "UList_41" : UInt = PLC HMI_IF.UList[41] AT %DB1.DBW0, 100 ms   // HMI_IF.UList[41]
   "UList_42" : UInt = PLC HMI_IF.UList[42] AT %DB1.DBW0, 100 ms   // HMI_IF.UList[42]
   "UList_43" : UInt = PLC HMI_IF.UList[43] AT %DB1.DBW0, 100 ms   // HMI_IF.UList[43]
   "UList_44" : UInt = PLC HMI_IF.UList[44] AT %DB1.DBW0, 100 ms   // HMI_IF.UList[44]
   "UList_45" : UInt = PLC HMI_IF.UList[45] AT %DB1.DBW0, 100 ms   // HMI_IF.UList[45]
   "UList_46" : UInt = PLC HMI_IF.UList[46] AT %DB1.DBW0, 100 ms   // HMI_IF.UList[46]
   "UList_47" : UInt = PLC HMI_IF.UList[47] AT %DB1.DBW0, 100 ms   // HMI_IF.UList[47]
   "UList_48" : UInt = PLC HMI_IF.UList[48] AT %DB1.DBW0, 100 ms   // HMI_IF.UList[48]
   "LList_01" : UInt = PLC HMI_IF.LList[1] AT %DB1.DBW0, 100 ms   // HMI_IF.LList[1]
   "LList_02" : UInt = PLC HMI_IF.LList[2] AT %DB1.DBW0, 100 ms   // HMI_IF.LList[2]
   "LList_03" : UInt = PLC HMI_IF.LList[3] AT %DB1.DBW0, 100 ms   // HMI_IF.LList[3]
   "LList_04" : UInt = PLC HMI_IF.LList[4] AT %DB1.DBW0, 100 ms   // HMI_IF.LList[4]
   "LList_05" : UInt = PLC HMI_IF.LList[5] AT %DB1.DBW0, 100 ms   // HMI_IF.LList[5]
   "LList_06" : UInt = PLC HMI_IF.LList[6] AT %DB1.DBW0, 100 ms   // HMI_IF.LList[6]
   "LList_07" : UInt = PLC HMI_IF.LList[7] AT %DB1.DBW0, 100 ms   // HMI_IF.LList[7]
   "LList_08" : UInt = PLC HMI_IF.LList[8] AT %DB1.DBW0, 100 ms   // HMI_IF.LList[8]
   "LList_09" : UInt = PLC HMI_IF.LList[9] AT %DB1.DBW0, 100 ms   // HMI_IF.LList[9]
   "LList_10" : UInt = PLC HMI_IF.LList[10] AT %DB1.DBW0, 100 ms   // HMI_IF.LList[10]
   "LList_11" : UInt = PLC HMI_IF.LList[11] AT %DB1.DBW0, 100 ms   // HMI_IF.LList[11]
   "LList_12" : UInt = PLC HMI_IF.LList[12] AT %DB1.DBW0, 100 ms   // HMI_IF.LList[12]
   "LList_13" : UInt = PLC HMI_IF.LList[13] AT %DB1.DBW0, 100 ms   // HMI_IF.LList[13]
   "LList_14" : UInt = PLC HMI_IF.LList[14] AT %DB1.DBW0, 100 ms   // HMI_IF.LList[14]
   "LList_15" : UInt = PLC HMI_IF.LList[15] AT %DB1.DBW0, 100 ms   // HMI_IF.LList[15]
   "LList_16" : UInt = PLC HMI_IF.LList[16] AT %DB1.DBW0, 100 ms   // HMI_IF.LList[16]
   "LList_17" : UInt = PLC HMI_IF.LList[17] AT %DB1.DBW0, 100 ms   // HMI_IF.LList[17]
   "LList_18" : UInt = PLC HMI_IF.LList[18] AT %DB1.DBW0, 100 ms   // HMI_IF.LList[18]
   "LList_19" : UInt = PLC HMI_IF.LList[19] AT %DB1.DBW0, 100 ms   // HMI_IF.LList[19]
   "LList_20" : UInt = PLC HMI_IF.LList[20] AT %DB1.DBW0, 100 ms   // HMI_IF.LList[20]
   "LList_21" : UInt = PLC HMI_IF.LList[21] AT %DB1.DBW0, 100 ms   // HMI_IF.LList[21]
   "LList_22" : UInt = PLC HMI_IF.LList[22] AT %DB1.DBW0, 100 ms   // HMI_IF.LList[22]
   "LList_23" : UInt = PLC HMI_IF.LList[23] AT %DB1.DBW0, 100 ms   // HMI_IF.LList[23]
   "LList_24" : UInt = PLC HMI_IF.LList[24] AT %DB1.DBW0, 100 ms   // HMI_IF.LList[24]
   "LList_25" : UInt = PLC HMI_IF.LList[25] AT %DB1.DBW0, 100 ms   // HMI_IF.LList[25]
   "LList_26" : UInt = PLC HMI_IF.LList[26] AT %DB1.DBW0, 100 ms   // HMI_IF.LList[26]
   "LList_27" : UInt = PLC HMI_IF.LList[27] AT %DB1.DBW0, 100 ms   // HMI_IF.LList[27]
   "LList_28" : UInt = PLC HMI_IF.LList[28] AT %DB1.DBW0, 100 ms   // HMI_IF.LList[28]
   "LList_29" : UInt = PLC HMI_IF.LList[29] AT %DB1.DBW0, 100 ms   // HMI_IF.LList[29]
   "LList_30" : UInt = PLC HMI_IF.LList[30] AT %DB1.DBW0, 100 ms   // HMI_IF.LList[30]
   "LList_31" : UInt = PLC HMI_IF.LList[31] AT %DB1.DBW0, 100 ms   // HMI_IF.LList[31]
   "LList_32" : UInt = PLC HMI_IF.LList[32] AT %DB1.DBW0, 100 ms   // HMI_IF.LList[32]
   "LList_33" : UInt = PLC HMI_IF.LList[33] AT %DB1.DBW0, 100 ms   // HMI_IF.LList[33]
   "LList_34" : UInt = PLC HMI_IF.LList[34] AT %DB1.DBW0, 100 ms   // HMI_IF.LList[34]
   "LList_35" : UInt = PLC HMI_IF.LList[35] AT %DB1.DBW0, 100 ms   // HMI_IF.LList[35]
   "LList_36" : UInt = PLC HMI_IF.LList[36] AT %DB1.DBW0, 100 ms   // HMI_IF.LList[36]
   "LList_37" : UInt = PLC HMI_IF.LList[37] AT %DB1.DBW0, 100 ms   // HMI_IF.LList[37]
   "LList_38" : UInt = PLC HMI_IF.LList[38] AT %DB1.DBW0, 100 ms   // HMI_IF.LList[38]
   "LList_39" : UInt = PLC HMI_IF.LList[39] AT %DB1.DBW0, 100 ms   // HMI_IF.LList[39]
   "LList_40" : UInt = PLC HMI_IF.LList[40] AT %DB1.DBW0, 100 ms   // HMI_IF.LList[40]
   "LList_41" : UInt = PLC HMI_IF.LList[41] AT %DB1.DBW0, 100 ms   // HMI_IF.LList[41]
   "LList_42" : UInt = PLC HMI_IF.LList[42] AT %DB1.DBW0, 100 ms   // HMI_IF.LList[42]
   "LList_43" : UInt = PLC HMI_IF.LList[43] AT %DB1.DBW0, 100 ms   // HMI_IF.LList[43]
   "LList_44" : UInt = PLC HMI_IF.LList[44] AT %DB1.DBW0, 100 ms   // HMI_IF.LList[44]
   "LList_45" : UInt = PLC HMI_IF.LList[45] AT %DB1.DBW0, 100 ms   // HMI_IF.LList[45]
   "LList_46" : UInt = PLC HMI_IF.LList[46] AT %DB1.DBW0, 100 ms   // HMI_IF.LList[46]
   "LList_47" : UInt = PLC HMI_IF.LList[47] AT %DB1.DBW0, 100 ms   // HMI_IF.LList[47]
   "LList_48" : UInt = PLC HMI_IF.LList[48] AT %DB1.DBW0, 100 ms   // HMI_IF.LList[48]
   "UState_01" : USInt = PLC HMI_IF.UState[1] AT %DB1.DBW0, 100 ms   // HMI_IF.UState[1]
   "UState_02" : USInt = PLC HMI_IF.UState[2] AT %DB1.DBW0, 100 ms   // HMI_IF.UState[2]
   "UState_03" : USInt = PLC HMI_IF.UState[3] AT %DB1.DBW0, 100 ms   // HMI_IF.UState[3]
   "UState_04" : USInt = PLC HMI_IF.UState[4] AT %DB1.DBW0, 100 ms   // HMI_IF.UState[4]
   "UState_05" : USInt = PLC HMI_IF.UState[5] AT %DB1.DBW0, 100 ms   // HMI_IF.UState[5]
   "UState_06" : USInt = PLC HMI_IF.UState[6] AT %DB1.DBW0, 100 ms   // HMI_IF.UState[6]
   "UState_07" : USInt = PLC HMI_IF.UState[7] AT %DB1.DBW0, 100 ms   // HMI_IF.UState[7]
   "UState_08" : USInt = PLC HMI_IF.UState[8] AT %DB1.DBW0, 100 ms   // HMI_IF.UState[8]
   "UState_09" : USInt = PLC HMI_IF.UState[9] AT %DB1.DBW0, 100 ms   // HMI_IF.UState[9]
   "UState_10" : USInt = PLC HMI_IF.UState[10] AT %DB1.DBW0, 100 ms   // HMI_IF.UState[10]
   "UState_11" : USInt = PLC HMI_IF.UState[11] AT %DB1.DBW0, 100 ms   // HMI_IF.UState[11]
   "UState_12" : USInt = PLC HMI_IF.UState[12] AT %DB1.DBW0, 100 ms   // HMI_IF.UState[12]
   "UState_13" : USInt = PLC HMI_IF.UState[13] AT %DB1.DBW0, 100 ms   // HMI_IF.UState[13]
   "UState_14" : USInt = PLC HMI_IF.UState[14] AT %DB1.DBW0, 100 ms   // HMI_IF.UState[14]
   "UState_15" : USInt = PLC HMI_IF.UState[15] AT %DB1.DBW0, 100 ms   // HMI_IF.UState[15]
   "UState_16" : USInt = PLC HMI_IF.UState[16] AT %DB1.DBW0, 100 ms   // HMI_IF.UState[16]
   "UState_17" : USInt = PLC HMI_IF.UState[17] AT %DB1.DBW0, 100 ms   // HMI_IF.UState[17]
   "UState_18" : USInt = PLC HMI_IF.UState[18] AT %DB1.DBW0, 100 ms   // HMI_IF.UState[18]
   "UState_19" : USInt = PLC HMI_IF.UState[19] AT %DB1.DBW0, 100 ms   // HMI_IF.UState[19]
   "UState_20" : USInt = PLC HMI_IF.UState[20] AT %DB1.DBW0, 100 ms   // HMI_IF.UState[20]
   "UState_21" : USInt = PLC HMI_IF.UState[21] AT %DB1.DBW0, 100 ms   // HMI_IF.UState[21]
   "UState_22" : USInt = PLC HMI_IF.UState[22] AT %DB1.DBW0, 100 ms   // HMI_IF.UState[22]
   "UState_23" : USInt = PLC HMI_IF.UState[23] AT %DB1.DBW0, 100 ms   // HMI_IF.UState[23]
   "UState_24" : USInt = PLC HMI_IF.UState[24] AT %DB1.DBW0, 100 ms   // HMI_IF.UState[24]
   "UState_25" : USInt = PLC HMI_IF.UState[25] AT %DB1.DBW0, 100 ms   // HMI_IF.UState[25]
   "UState_26" : USInt = PLC HMI_IF.UState[26] AT %DB1.DBW0, 100 ms   // HMI_IF.UState[26]
   "UState_27" : USInt = PLC HMI_IF.UState[27] AT %DB1.DBW0, 100 ms   // HMI_IF.UState[27]
   "UState_28" : USInt = PLC HMI_IF.UState[28] AT %DB1.DBW0, 100 ms   // HMI_IF.UState[28]
   "UState_29" : USInt = PLC HMI_IF.UState[29] AT %DB1.DBW0, 100 ms   // HMI_IF.UState[29]
   "UState_30" : USInt = PLC HMI_IF.UState[30] AT %DB1.DBW0, 100 ms   // HMI_IF.UState[30]
   "UState_31" : USInt = PLC HMI_IF.UState[31] AT %DB1.DBW0, 100 ms   // HMI_IF.UState[31]
   "UState_32" : USInt = PLC HMI_IF.UState[32] AT %DB1.DBW0, 100 ms   // HMI_IF.UState[32]
   "UState_33" : USInt = PLC HMI_IF.UState[33] AT %DB1.DBW0, 100 ms   // HMI_IF.UState[33]
   "UState_34" : USInt = PLC HMI_IF.UState[34] AT %DB1.DBW0, 100 ms   // HMI_IF.UState[34]
   "UState_35" : USInt = PLC HMI_IF.UState[35] AT %DB1.DBW0, 100 ms   // HMI_IF.UState[35]
   "UState_36" : USInt = PLC HMI_IF.UState[36] AT %DB1.DBW0, 100 ms   // HMI_IF.UState[36]
   "UState_37" : USInt = PLC HMI_IF.UState[37] AT %DB1.DBW0, 100 ms   // HMI_IF.UState[37]
   "UState_38" : USInt = PLC HMI_IF.UState[38] AT %DB1.DBW0, 100 ms   // HMI_IF.UState[38]
   "UState_39" : USInt = PLC HMI_IF.UState[39] AT %DB1.DBW0, 100 ms   // HMI_IF.UState[39]
   "UState_40" : USInt = PLC HMI_IF.UState[40] AT %DB1.DBW0, 100 ms   // HMI_IF.UState[40]
   "UState_41" : USInt = PLC HMI_IF.UState[41] AT %DB1.DBW0, 100 ms   // HMI_IF.UState[41]
   "UState_42" : USInt = PLC HMI_IF.UState[42] AT %DB1.DBW0, 100 ms   // HMI_IF.UState[42]
   "UState_43" : USInt = PLC HMI_IF.UState[43] AT %DB1.DBW0, 100 ms   // HMI_IF.UState[43]
   "UState_44" : USInt = PLC HMI_IF.UState[44] AT %DB1.DBW0, 100 ms   // HMI_IF.UState[44]
   "UState_45" : USInt = PLC HMI_IF.UState[45] AT %DB1.DBW0, 100 ms   // HMI_IF.UState[45]
   "UState_46" : USInt = PLC HMI_IF.UState[46] AT %DB1.DBW0, 100 ms   // HMI_IF.UState[46]
   "UState_47" : USInt = PLC HMI_IF.UState[47] AT %DB1.DBW0, 100 ms   // HMI_IF.UState[47]
   "UState_48" : USInt = PLC HMI_IF.UState[48] AT %DB1.DBW0, 100 ms   // HMI_IF.UState[48]
   "LState_01" : USInt = PLC HMI_IF.LState[1] AT %DB1.DBW0, 100 ms   // HMI_IF.LState[1]
   "LState_02" : USInt = PLC HMI_IF.LState[2] AT %DB1.DBW0, 100 ms   // HMI_IF.LState[2]
   "LState_03" : USInt = PLC HMI_IF.LState[3] AT %DB1.DBW0, 100 ms   // HMI_IF.LState[3]
   "LState_04" : USInt = PLC HMI_IF.LState[4] AT %DB1.DBW0, 100 ms   // HMI_IF.LState[4]
   "LState_05" : USInt = PLC HMI_IF.LState[5] AT %DB1.DBW0, 100 ms   // HMI_IF.LState[5]
   "LState_06" : USInt = PLC HMI_IF.LState[6] AT %DB1.DBW0, 100 ms   // HMI_IF.LState[6]
   "LState_07" : USInt = PLC HMI_IF.LState[7] AT %DB1.DBW0, 100 ms   // HMI_IF.LState[7]
   "LState_08" : USInt = PLC HMI_IF.LState[8] AT %DB1.DBW0, 100 ms   // HMI_IF.LState[8]
   "LState_09" : USInt = PLC HMI_IF.LState[9] AT %DB1.DBW0, 100 ms   // HMI_IF.LState[9]
   "LState_10" : USInt = PLC HMI_IF.LState[10] AT %DB1.DBW0, 100 ms   // HMI_IF.LState[10]
   "LState_11" : USInt = PLC HMI_IF.LState[11] AT %DB1.DBW0, 100 ms   // HMI_IF.LState[11]
   "LState_12" : USInt = PLC HMI_IF.LState[12] AT %DB1.DBW0, 100 ms   // HMI_IF.LState[12]
   "LState_13" : USInt = PLC HMI_IF.LState[13] AT %DB1.DBW0, 100 ms   // HMI_IF.LState[13]
   "LState_14" : USInt = PLC HMI_IF.LState[14] AT %DB1.DBW0, 100 ms   // HMI_IF.LState[14]
   "LState_15" : USInt = PLC HMI_IF.LState[15] AT %DB1.DBW0, 100 ms   // HMI_IF.LState[15]
   "LState_16" : USInt = PLC HMI_IF.LState[16] AT %DB1.DBW0, 100 ms   // HMI_IF.LState[16]
   "LState_17" : USInt = PLC HMI_IF.LState[17] AT %DB1.DBW0, 100 ms   // HMI_IF.LState[17]
   "LState_18" : USInt = PLC HMI_IF.LState[18] AT %DB1.DBW0, 100 ms   // HMI_IF.LState[18]
   "LState_19" : USInt = PLC HMI_IF.LState[19] AT %DB1.DBW0, 100 ms   // HMI_IF.LState[19]
   "LState_20" : USInt = PLC HMI_IF.LState[20] AT %DB1.DBW0, 100 ms   // HMI_IF.LState[20]
   "LState_21" : USInt = PLC HMI_IF.LState[21] AT %DB1.DBW0, 100 ms   // HMI_IF.LState[21]
   "LState_22" : USInt = PLC HMI_IF.LState[22] AT %DB1.DBW0, 100 ms   // HMI_IF.LState[22]
   "LState_23" : USInt = PLC HMI_IF.LState[23] AT %DB1.DBW0, 100 ms   // HMI_IF.LState[23]
   "LState_24" : USInt = PLC HMI_IF.LState[24] AT %DB1.DBW0, 100 ms   // HMI_IF.LState[24]
   "LState_25" : USInt = PLC HMI_IF.LState[25] AT %DB1.DBW0, 100 ms   // HMI_IF.LState[25]
   "LState_26" : USInt = PLC HMI_IF.LState[26] AT %DB1.DBW0, 100 ms   // HMI_IF.LState[26]
   "LState_27" : USInt = PLC HMI_IF.LState[27] AT %DB1.DBW0, 100 ms   // HMI_IF.LState[27]
   "LState_28" : USInt = PLC HMI_IF.LState[28] AT %DB1.DBW0, 100 ms   // HMI_IF.LState[28]
   "LState_29" : USInt = PLC HMI_IF.LState[29] AT %DB1.DBW0, 100 ms   // HMI_IF.LState[29]
   "LState_30" : USInt = PLC HMI_IF.LState[30] AT %DB1.DBW0, 100 ms   // HMI_IF.LState[30]
   "LState_31" : USInt = PLC HMI_IF.LState[31] AT %DB1.DBW0, 100 ms   // HMI_IF.LState[31]
   "LState_32" : USInt = PLC HMI_IF.LState[32] AT %DB1.DBW0, 100 ms   // HMI_IF.LState[32]
   "LState_33" : USInt = PLC HMI_IF.LState[33] AT %DB1.DBW0, 100 ms   // HMI_IF.LState[33]
   "LState_34" : USInt = PLC HMI_IF.LState[34] AT %DB1.DBW0, 100 ms   // HMI_IF.LState[34]
   "LState_35" : USInt = PLC HMI_IF.LState[35] AT %DB1.DBW0, 100 ms   // HMI_IF.LState[35]
   "LState_36" : USInt = PLC HMI_IF.LState[36] AT %DB1.DBW0, 100 ms   // HMI_IF.LState[36]
   "LState_37" : USInt = PLC HMI_IF.LState[37] AT %DB1.DBW0, 100 ms   // HMI_IF.LState[37]
   "LState_38" : USInt = PLC HMI_IF.LState[38] AT %DB1.DBW0, 100 ms   // HMI_IF.LState[38]
   "LState_39" : USInt = PLC HMI_IF.LState[39] AT %DB1.DBW0, 100 ms   // HMI_IF.LState[39]
   "LState_40" : USInt = PLC HMI_IF.LState[40] AT %DB1.DBW0, 100 ms   // HMI_IF.LState[40]
   "LState_41" : USInt = PLC HMI_IF.LState[41] AT %DB1.DBW0, 100 ms   // HMI_IF.LState[41]
   "LState_42" : USInt = PLC HMI_IF.LState[42] AT %DB1.DBW0, 100 ms   // HMI_IF.LState[42]
   "LState_43" : USInt = PLC HMI_IF.LState[43] AT %DB1.DBW0, 100 ms   // HMI_IF.LState[43]
   "LState_44" : USInt = PLC HMI_IF.LState[44] AT %DB1.DBW0, 100 ms   // HMI_IF.LState[44]
   "LState_45" : USInt = PLC HMI_IF.LState[45] AT %DB1.DBW0, 100 ms   // HMI_IF.LState[45]
   "LState_46" : USInt = PLC HMI_IF.LState[46] AT %DB1.DBW0, 100 ms   // HMI_IF.LState[46]
   "LState_47" : USInt = PLC HMI_IF.LState[47] AT %DB1.DBW0, 100 ms   // HMI_IF.LState[47]
   "LState_48" : USInt = PLC HMI_IF.LState[48] AT %DB1.DBW0, 100 ms   // HMI_IF.LState[48]
   "BalL" : Int = PLC HMI_IF.BalL AT %DB1.DBW0, 100 ms   // HMI_IF.BalL
   "BalR" : Int = PLC HMI_IF.BalR AT %DB1.DBW0, 100 ms   // HMI_IF.BalR
   "BalDiff" : Int = PLC HMI_IF.BalDiff AT %DB1.DBW0, 100 ms   // HMI_IF.BalDiff
   "BalF" : Int = PLC HMI_IF.BalF AT %DB1.DBW0, 100 ms   // HMI_IF.BalF
   "BalA" : Int = PLC HMI_IF.BalA AT %DB1.DBW0, 100 ms   // HMI_IF.BalA
   "BalOk" : Bool = PLC HMI_IF.BalOk AT %DB1.DBW0, 100 ms   // HMI_IF.BalOk
   "AlarmWord" : Word = PLC HMI_IF.AlarmWord AT %DB1.DBW0, 100 ms   // HMI_IF.AlarmWord
   "AlarmAckWord" : Word = PLC HMI_IF.AlarmAckWord AT %DB1.DBW0, 100 ms   // HMI_IF.AlarmAckWord
   "AlarmId" : UInt = PLC HMI_IF.AlarmId AT %DB1.DBW0, 100 ms   // HMI_IF.AlarmId
   "AlarmWord2" : Word = PLC HMI_IF.AlarmWord2 AT %DB1.DBW0, 100 ms   // HMI_IF.AlarmWord2
   "AlarmUId" : UInt = PLC HMI_IF.AlarmUId AT %DB1.DBW0, 100 ms   // HMI_IF.AlarmUId
   "AlarmUCnt" : Int = PLC HMI_IF.AlarmUCnt AT %DB1.DBW0, 100 ms   // HMI_IF.AlarmUCnt
   "AlarmLId" : UInt = PLC HMI_IF.AlarmLId AT %DB1.DBW0, 100 ms   // HMI_IF.AlarmLId
   "AlarmLCnt" : Int = PLC HMI_IF.AlarmLCnt AT %DB1.DBW0, 100 ms   // HMI_IF.AlarmLCnt
   "AlarmX" : SInt = PLC HMI_IF.AlarmX AT %DB1.DBW0, 100 ms   // HMI_IF.AlarmX
   "AlarmY" : SInt = PLC HMI_IF.AlarmY AT %DB1.DBW0, 100 ms   // HMI_IF.AlarmY
   "AlarmBay" : USInt = PLC HMI_IF.AlarmBay AT %DB1.DBW0, 100 ms   // HMI_IF.AlarmBay
   "AlarmHist_00" : Int = PLC HMI_IF.AlarmHist[0] AT %DB1.DBW0, 100 ms   // HMI_IF.AlarmHist[0]
   "AlarmHist_01" : Int = PLC HMI_IF.AlarmHist[1] AT %DB1.DBW0, 100 ms   // HMI_IF.AlarmHist[1]
   "AlarmHist_02" : Int = PLC HMI_IF.AlarmHist[2] AT %DB1.DBW0, 100 ms   // HMI_IF.AlarmHist[2]
   "AlarmHist_03" : Int = PLC HMI_IF.AlarmHist[3] AT %DB1.DBW0, 100 ms   // HMI_IF.AlarmHist[3]
   "AlarmHist_04" : Int = PLC HMI_IF.AlarmHist[4] AT %DB1.DBW0, 100 ms   // HMI_IF.AlarmHist[4]
   "AlarmHist_05" : Int = PLC HMI_IF.AlarmHist[5] AT %DB1.DBW0, 100 ms   // HMI_IF.AlarmHist[5]
   "AlarmHist_06" : Int = PLC HMI_IF.AlarmHist[6] AT %DB1.DBW0, 100 ms   // HMI_IF.AlarmHist[6]
   "AlarmHist_07" : Int = PLC HMI_IF.AlarmHist[7] AT %DB1.DBW0, 100 ms   // HMI_IF.AlarmHist[7]
   "AlarmHist_08" : Int = PLC HMI_IF.AlarmHist[8] AT %DB1.DBW0, 100 ms   // HMI_IF.AlarmHist[8]
   "AlarmHist_09" : Int = PLC HMI_IF.AlarmHist[9] AT %DB1.DBW0, 100 ms   // HMI_IF.AlarmHist[9]
   "AlarmHist_10" : Int = PLC HMI_IF.AlarmHist[10] AT %DB1.DBW0, 100 ms   // HMI_IF.AlarmHist[10]
   "AlarmHist_11" : Int = PLC HMI_IF.AlarmHist[11] AT %DB1.DBW0, 100 ms   // HMI_IF.AlarmHist[11]
   "AlarmHist_12" : Int = PLC HMI_IF.AlarmHist[12] AT %DB1.DBW0, 100 ms   // HMI_IF.AlarmHist[12]
   "AlarmHist_13" : Int = PLC HMI_IF.AlarmHist[13] AT %DB1.DBW0, 100 ms   // HMI_IF.AlarmHist[13]
   "AlarmHist_14" : Int = PLC HMI_IF.AlarmHist[14] AT %DB1.DBW0, 100 ms   // HMI_IF.AlarmHist[14]
   "AlarmHist_15" : Int = PLC HMI_IF.AlarmHist[15] AT %DB1.DBW0, 100 ms   // HMI_IF.AlarmHist[15]
   "AlarmHistSeq" : UDInt = PLC HMI_IF.AlarmHistSeq AT %DB1.DBW0, 100 ms   // HMI_IF.AlarmHistSeq
   "OB30Ticks" : UDInt = PLC HMI_IF.OB30Ticks AT %DB1.DBW0, 100 ms   // HMI_IF.OB30Ticks
   "Heartbeat" : Bool = PLC HMI_IF.Heartbeat AT %DB1.DBW0, 100 ms   // HMI_IF.Heartbeat

discrete alarms
   1: 'EN: Ship imbalance |L-R| > 5. Blokirajući: DA iz OB30 provjere, inače upozorenje. Bit 0 u HMI_IF.AlarmWord. / Neuravnoteženost broda: razlika lijeve i desne polovice > 5', class Errors, trigger "AlarmWord" bit 0
   2: 'EN: Pick location empty. Blokirajući: DA. Bit 1 u HMI_IF.AlarmWord. / Lokacija s koje se podiže kontejner je prazna', class Errors, trigger "AlarmWord" bit 1
   3: 'EN: Drop location occupied. Blokirajući: DA. Bit 2 u HMI_IF.AlarmWord. / Lokacija na koju se spušta kontejner je zauzeta', class Errors, trigger "AlarmWord" bit 2
   4: 'EN: Unload ID not in Bay 0. Blokirajući: NE. Bit 3 u HMI_IF.AlarmWord. / ID kontejnera postoji u listi za istovar, ali ne postoji u polju Bay 0', class Warnings, trigger "AlarmWord" bit 3
   5: 'EN: Load ID not in Bay 1. Blokirajući: NE. Bit 4 u HMI_IF.AlarmWord. / ID kontejnera postoji u listi za ukrcaj, ali ne postoji u polju Bay 1', class Warnings, trigger "AlarmWord" bit 4
   6: 'EN: Invalid container ID. Blokirajući: NE. Bit 5 u HMI_IF.AlarmWord. / Neispravan ID kontejnera (izvan 100–999)', class Warnings, trigger "AlarmWord" bit 5
   7: 'EN: Duplicate container ID. Blokirajući: NE. Bit 6 u HMI_IF.AlarmWord. / Dvostruki ID kontejnera', class Warnings, trigger "AlarmWord" bit 6
   8: 'EN: No free slot. Blokirajući: DA. Bit 7 u HMI_IF.AlarmWord. / Nema slobodnog mjesta u odredišnom polju', class Errors, trigger "AlarmWord" bit 7
   9: 'EN: Plan infeasible. Blokirajući: DA. Bit 8 u HMI_IF.AlarmWord. / Plan istovara/ukrcaja nije izvediv', class Errors, trigger "AlarmWord" bit 8
   10: 'EN: Invalid manual command. Blokirajući: DA iz OB30 provjere, inače upozorenje. Bit 9 u HMI_IF.AlarmWord. / Neispravna ručna naredba (Bay mora biti 0/1, x 0–3, y 0–11)', class Errors, trigger "AlarmWord" bit 9
   11: 'EN: FB1 timeout. Blokirajući: DA. Bit 10 u HMI_IF.AlarmWord. / Dizalica nije izvršila naredbu (timeout)', class Errors, trigger "AlarmWord" bit 10
   12: 'EN: Crane already carrying. Blokirajući: DA. Bit 11 u HMI_IF.AlarmWord. / Dizalica već nosi kontejner', class Errors, trigger "AlarmWord" bit 11
   13: 'EN: Crane is empty (put down). Blokirajući: DA. Bit 12 u HMI_IF.AlarmWord. / Dizalica ne nosi kontejner', class Errors, trigger "AlarmWord" bit 12
   14: 'EN: Not initialized. Blokirajući: NE. Bit 13 u HMI_IF.AlarmWord. / Sustav nije inicijaliziran: pritisnite POČETNO STANJE', class Warnings, trigger "AlarmWord" bit 13
   15: 'EN: Crane position mismatch after move. Blokirajući: DA. Bit 14 u HMI_IF.AlarmWord. / Položaj dizalice ne odgovara naredbi', class Errors, trigger "AlarmWord" bit 14
   16: 'EN: Unloading and loading finished. Blokirajući: NE. Bit 15 u HMI_IF.AlarmWord. / Istovar i ukrcaj završeni', class Warnings, trigger "AlarmWord" bit 15
   17: 'EN: List order infeasible under the balance rule: plan uses free order. Blokirajući: NE. Bit 0 u HMI_IF.AlarmWord2. / Liste se ne mogu izvršiti zadanim redoslijedom zbog ravnoteže broda: plan koristi slobodan redoslijed', class Warnings, trigger "AlarmWord2" bit 0
   18: 'EN: Ship loaded out of balance: plan keeps the list order, |L-R| never exceeds the start value and ends <= 5. Blokirajući: NE. Bit 1 u HMI_IF.AlarmWord2. / Brod je zadan neuravnotežen: plan drži zadani redoslijed, |L-D| ne prelazi početnu razliku i završava <= 5', class Warnings, trigger "AlarmWord2" bit 1

text list "TL_Alarm": -1 '-'; 0 '0 Neuravnoteženost broda |L-R| > 5'; 1 '1 Lokacija podizanja prazna'; 2 '2 Lokacija spuštanja zauzeta'; 3 '3 ID u listi za istovar, nije u Bay 0'; 4 '4 ID u listi za ukrcaj, nije u Bay 1'; 5 '5 Neispravan ID (100-999)'; 6 '6 Dvostruki ID'; 7 '7 Nema slobodnog mjesta'; 8 '8 Plan nije izvediv'; 9 '9 Neispravna ručna naredba'; 10 '10 Dizalica: timeout naredbe'; 11 '11 Dizalica već nosi kontejner'; 12 '12 Dizalica ne nosi kontejner'; 13 '13 Nije inicijalizirano'; 14 '14 Položaj dizalice ne odgovara'; 15 '15 Istovar i ukrcaj završeni'

text list "TL_BalMode": 0 '0 lijevo/desno'; 1 '1 + pramac/krma'

text list "TL_Bay": 0 '0 BROD'; 1 '1 SKLADIŠTE'

text list "TL_Cmd": 0 '-'; 1 '1 PODIGNI'; 2 '2 SPUSTI'; 3 '3 POMAKNI'; 10 '10 RESET'

text list "TL_Kind": 0 '-'; 1 'ISTOVAR Bay0->Bay1'; 2 'UKRCAJ Bay1->Bay0'

text list "TL_ListSt": 0 'čeka'; 1 'gotovo'; 2 'preskočeno'; 3 'u tijeku'

text list "TL_Mode": 0 '-'; 1 'AUTOMATSKI'; 2 'POLUAUTOMATSKI'; 3 'RUČNO'

text list "TL_Order": 0 '0 slobodan redoslijed'; 1 '1 redoslijed po listi'; 2 '2 strogo: istovar pa ukrcaj'

text list "TL_Phase": 0 'vožnja do izvora'; 1 'podizanje'; 2 'vožnja do odredišta'; 3 'spuštanje'

text list "TL_State": 0 'ISKLJUČENO'; 1 'INICIJALIZACIJA'; 2 'SPREMAN'; 3 'RADI'; 4 'PAUZA'; 5 'ALARM'; 6 'ZAVRŠENO'; 7 'PLANIRANJE'

text list "TL_YesNo": 0 'NE'; 1 'DA'

screen "Alarms" 1920x1080, template "Tpl"
   AlarmView "Alarm view_1" at 16,190 size 1580x300
   AlarmView "Alarm view_2" at 16,600 size 1580x350
   TextField "Text field_1" at 26,153 size 134x22; Text 'AKTIVNI ALARMI'
   TextField "Text field_2" at 26,563 size 147x22; Text 'POVIJEST ALARMA'

Template "Tpl" 1920x1080
   TextField "hdr_frm_1" at 0,0 size 1920x148; Text 'Text'
   TextField "hdr_txt_1" at 16,10 size 270x34; Text 'LUČKA DIZALICA'
   TextField "hdr_txt_2" at 16,44 size 270x22; Text 'PLC Challenge 2026 - EESTEC'
   Rectangle "hdr_lmp_1" at 290,14 size 14x14
      Appearance <- "Heartbeat"
   Button "hdr_btn_1" at 320,10 size 160x58; TextOff 'UKLJ. / ISKLJ.'
      on Press: InvertBit("SwOn")
   Rectangle "hdr_lmp_2" at 490,12 size 22x22
      Appearance <- "LampReady"
   TextField "hdr_txt_3" at 516,12 size 110x22; Text 'SPREMAN'
   Rectangle "hdr_lmp_3" at 490,44 size 22x22
      Appearance <- "LampOff"
   TextField "hdr_txt_4" at 516,44 size 110x22; Text 'ISKLJ.'
   Button "hdr_btn_2" at 640,10 size 180x58; TextOff 'INIT'
      on Press: SetBit("BtnInit")
   Button "hdr_btn_3" at 840,10 size 160x58; TextOff 'AUTO'
      on Press: SetBit("BtnAuto")
   Rectangle "hdr_lmp_4" at 840,70 size 160x8
      Appearance <- "LampAuto"
   Button "hdr_btn_4" at 1006,10 size 180x58; TextOff 'SEMI'
      on Press: SetBit("BtnSemi")
   Rectangle "hdr_lmp_5" at 1006,70 size 180x8
      Appearance <- "LampSemi"
   Button "hdr_btn_5" at 1192,10 size 140x58; TextOff 'RUČNO'
      on Press: SetBit("BtnManual")
   Rectangle "hdr_lmp_6" at 1192,70 size 140x8
      Appearance <- "LampManual"
   Button "hdr_btn_6" at 1352,10 size 120x58; TextOff 'START'
      on Press: SetBit("BtnStart")
   Rectangle "hdr_lmp_7" at 1352,70 size 120x8
      Appearance <- "LampRunning"
   Button "hdr_btn_7" at 1478,10 size 120x58; TextOff 'STOP'
      on Press: SetBit("BtnStop")
   Button "hdr_btn_8" at 1604,10 size 120x58; TextOff 'POTVRDA'
      on Press: SetBit("BtnAck")
   Button "hdr_btn_9" at 1730,10 size 176x58; TextOff 'KORAK'
      on Press: SetBit("BtnStep")
   Rectangle "hdr_lmp_8" at 1730,70 size 176x8
      Appearance <- "StepWaiting"
   TextField "hdr_txt_5" at 16,92 size 80x34; Text 'ST.'
   SymbolicIOField "hdr_sym_1" at 96,92 size 200x34; TextOff '0'; TextOn '1'; TextList "TL_State"
      ProcessValue <- "State"
   SymbolicIOField "hdr_sym_2" at 302,92 size 178x34; TextOff '0'; TextOn '1'; TextList "TL_Mode"
      ProcessValue <- "Mode"
   TextField "hdr_txt_6" at 490,92 size 36x34; Text 'M'
   IOField "hdr_io_1" at 526,92 size 90x34; FormatPattern 99999
      ProcessValue <- "M"
   TextField "hdr_txt_7" at 622,92 size 50x34; Text 'T/s'
   IOField "hdr_io_2" at 672,92 size 110x34; FormatPattern 999999.9
      ProcessValue <- "T"
   TextField "hdr_txt_8" at 790,92 size 26x34; Text 'J'
   IOField "hdr_io_3" at 816,92 size 90x34; FormatPattern 9.9999
      ProcessValue <- "J"
   TextField "hdr_txt_9" at 914,92 size 112x34; Text 'Plan'
   IOField "hdr_io_4" at 1026,92 size 80x34; FormatPattern 99999
      ProcessValue <- "PredM"
   IOField "hdr_io_5" at 1110,92 size 104x34; FormatPattern 999999.9
      ProcessValue <- "PredT"
   IOField "hdr_io_6" at 1218,92 size 84x34; FormatPattern 9.9999
      ProcessValue <- "PredJ"
   TextField "hdr_txt_10" at 1312,92 size 54x34; Text 'Pr.'
   IOField "hdr_io_7" at 1366,92 size 52x34; FormatPattern 999
      ProcessValue <- "TrDone"
   TextField "hdr_txt_11" at 1418,92 size 12x34; Text '/'
   IOField "hdr_io_8" at 1430,92 size 52x34; FormatPattern 999
      ProcessValue <- "TrTotal"
   Rectangle "hdr_lmp_9" at 1494,98 size 22x22
      Appearance <- "LampAlarm"
   SymbolicIOField "hdr_sym_3" at 1520,92 size 386x34; TextOff '0'; TextOn '1'; TextList "TL_Alarm"
      ProcessValue <- "AlarmHist_00"
   TextField "hdr_frm_2" at 0,1024 size 1920x56; Text 'Text'
   Button "hdr_nav_1" at 16,1030 size 200x44; TextOff 'PRIKAZ'
      on Press: ActivateScreen("Screen_1", 0)
   Button "hdr_nav_2" at 226,1030 size 200x44; TextOff 'RUČNO'
      on Press: ActivateScreen("Manual", 0)
   Button "hdr_nav_3" at 436,1030 size 200x44; TextOff 'POSTAVKE'
      on Press: ActivateScreen("Lists", 0)
   Button "hdr_nav_4" at 646,1030 size 200x44; TextOff 'ALARMI'
      on Press: ActivateScreen("Alarms", 0)
   Button "hdr_nav_5" at 856,1030 size 200x44; TextOff 'POVIJEST'
      on Press: ActivateScreen("AlarmLog", 0)
   Button "hdr_nav_6" at 1066,1030 size 220x44; TextOff 'REZULTATI'
      on Press: ActivateScreen("Score", 0)
   TextField "hdr_txt_12" at 1300,1034 size 110x34; Text 'PLC takt'
   IOField "hdr_io_9" at 1410,1034 size 110x34; FormatPattern 9999999
      ProcessValue <- "OB30Ticks"
   DateTimeField "hdr_dtm_1" at 1560,1032 size 346x40

screen "AlarmLog" 1920x1080, template "Tpl"
   TextField "txt_1" at 16,156 size 1000x30; Text 'ZADNJIH 16 ALARMA ([0] najnoviji). Vremenska povijest: ALARMI.'
   TextField "txt_2" at 16,200 size 60x38; Text '[0]'
   SymbolicIOField "sym_1" at 80,200 size 1036x38; TextOff '0'; TextOn '1'; TextList "TL_Alarm"
      ProcessValue <- "AlarmHist_00"
   TextField "txt_3" at 16,246 size 60x38; Text '[1]'
   SymbolicIOField "sym_2" at 80,246 size 1036x38; TextOff '0'; TextOn '1'; TextList "TL_Alarm"
      ProcessValue <- "AlarmHist_01"
   TextField "txt_4" at 16,292 size 60x38; Text '[2]'
   SymbolicIOField "sym_3" at 80,292 size 1036x38; TextOff '0'; TextOn '1'; TextList "TL_Alarm"
      ProcessValue <- "AlarmHist_02"
   TextField "txt_5" at 16,338 size 60x38; Text '[3]'
   SymbolicIOField "sym_4" at 80,338 size 1036x38; TextOff '0'; TextOn '1'; TextList "TL_Alarm"
      ProcessValue <- "AlarmHist_03"
   TextField "txt_6" at 16,384 size 60x38; Text '[4]'
   SymbolicIOField "sym_5" at 80,384 size 1036x38; TextOff '0'; TextOn '1'; TextList "TL_Alarm"
      ProcessValue <- "AlarmHist_04"
   TextField "txt_7" at 16,430 size 60x38; Text '[5]'
   SymbolicIOField "sym_6" at 80,430 size 1036x38; TextOff '0'; TextOn '1'; TextList "TL_Alarm"
      ProcessValue <- "AlarmHist_05"
   TextField "txt_8" at 16,476 size 60x38; Text '[6]'
   SymbolicIOField "sym_7" at 80,476 size 1036x38; TextOff '0'; TextOn '1'; TextList "TL_Alarm"
      ProcessValue <- "AlarmHist_06"
   TextField "txt_9" at 16,522 size 60x38; Text '[7]'
   SymbolicIOField "sym_8" at 80,522 size 1036x38; TextOff '0'; TextOn '1'; TextList "TL_Alarm"
      ProcessValue <- "AlarmHist_07"
   TextField "txt_10" at 16,568 size 60x38; Text '[8]'
   SymbolicIOField "sym_9" at 80,568 size 1036x38; TextOff '0'; TextOn '1'; TextList "TL_Alarm"
      ProcessValue <- "AlarmHist_08"
   TextField "txt_11" at 16,614 size 60x38; Text '[9]'
   SymbolicIOField "sym_10" at 80,614 size 1036x38; TextOff '0'; TextOn '1'; TextList "TL_Alarm"
      ProcessValue <- "AlarmHist_09"
   TextField "txt_12" at 16,660 size 60x38; Text '[10]'
   SymbolicIOField "sym_11" at 80,660 size 1036x38; TextOff '0'; TextOn '1'; TextList "TL_Alarm"
      ProcessValue <- "AlarmHist_10"
   TextField "txt_13" at 16,706 size 60x38; Text '[11]'
   SymbolicIOField "sym_12" at 80,706 size 1036x38; TextOff '0'; TextOn '1'; TextList "TL_Alarm"
      ProcessValue <- "AlarmHist_11"
   TextField "txt_14" at 16,752 size 60x38; Text '[12]'
   SymbolicIOField "sym_13" at 80,752 size 1036x38; TextOff '0'; TextOn '1'; TextList "TL_Alarm"
      ProcessValue <- "AlarmHist_12"
   TextField "txt_15" at 16,798 size 60x38; Text '[13]'
   SymbolicIOField "sym_14" at 80,798 size 1036x38; TextOff '0'; TextOn '1'; TextList "TL_Alarm"
      ProcessValue <- "AlarmHist_13"
   TextField "txt_16" at 16,844 size 60x38; Text '[14]'
   SymbolicIOField "sym_15" at 80,844 size 1036x38; TextOff '0'; TextOn '1'; TextList "TL_Alarm"
      ProcessValue <- "AlarmHist_14"
   TextField "txt_17" at 16,890 size 60x38; Text '[15]'
   SymbolicIOField "sym_16" at 80,890 size 1036x38; TextOff '0'; TextOn '1'; TextList "TL_Alarm"
      ProcessValue <- "AlarmHist_15"
   TextField "frm_1" at 1220,200 size 684x300; Text 'Text'
   TextField "txt_18" at 1232,206 size 600x28; Text 'NAJNOVIJI ALARM - DETALJI'
   Rectangle "lmp_1" at 1232,246 size 22x22
      Appearance <- "LampAlarm"
   TextField "txt_19" at 1262,240 size 150x34; Text 'Kontejner ID'
   IOField "io_1" at 1412,240 size 80x34; FormatPattern 999
      ProcessValue <- "AlarmId"
   TextField "txt_20" at 1232,284 size 120x34; Text 'Lokacija x'
   IOField "io_2" at 1352,284 size 50x34; FormatPattern s9
      ProcessValue <- "AlarmX"
   TextField "txt_21" at 1420,284 size 30x34; Text 'y'
   IOField "io_3" at 1450,284 size 50x34; FormatPattern s99
      ProcessValue <- "AlarmY"
   TextField "txt_22" at 1540,284 size 60x34; Text 'Bay'
   SymbolicIOField "sym_17" at 1600,284 size 240x34; TextOff '0'; TextOn '1'; TextList "TL_Bay"
      ProcessValue <- "AlarmBay"
   TextField "txt_23" at 1232,328 size 180x34; Text 'Riječ alarma'
   IOField "io_4" at 1412,328 size 100x34; FormatPattern 99999
      ProcessValue <- "AlarmWord"
   TextField "txt_24" at 1232,372 size 180x34; Text 'Broj pojava'
   IOField "io_5" at 1412,372 size 100x34; FormatPattern 999999
      ProcessValue <- "AlarmHistSeq"
   TextField "txt_25" at 1232,420 size 660x60; Text 'Uklonite uzrok alarma pa pritisnite POTVRDA.'
   TextField "frm_2" at 1220,516 size 684x236; Text 'Text'
   TextField "txt_26" at 1232,522 size 660x28; Text 'PROVJERA LISTA (POČETNO STANJE)'
   TextField "txt_27" at 1232,558 size 330x34; Text 'Istovar: prvi ID izvan broda'
   IOField "io_6" at 1562,558 size 80x34; FormatPattern 999
      ProcessValue <- "AlarmUId"
   TextField "txt_28" at 1660,558 size 90x34; Text 'ukupno'
   IOField "io_7" at 1750,558 size 60x34; FormatPattern 99
      ProcessValue <- "AlarmUCnt"
   TextField "txt_29" at 1232,600 size 330x34; Text 'Ukrcaj: prvi ID izvan skladista'
   IOField "io_8" at 1562,600 size 80x34; FormatPattern 999
      ProcessValue <- "AlarmLId"
   TextField "txt_30" at 1660,600 size 90x34; Text 'ukupno'
   IOField "io_9" at 1750,600 size 60x34; FormatPattern 99
      ProcessValue <- "AlarmLCnt"
   TextField "txt_31" at 1232,642 size 330x34; Text 'Redoslijed liste napušten'
   SymbolicIOField "sym_18" at 1562,642 size 100x34; TextOff '0'; TextOn '1'; TextList "TL_YesNo"
      ProcessValue <- "OrderFallback"
   TextField "txt_32" at 1232,684 size 330x34; Text 'Korišteni način redoslijeda'
   SymbolicIOField "sym_19" at 1562,684 size 300x34; TextOff '0'; TextOn '1'; TextList "TL_Order"
      ProcessValue <- "OrderModeAct"

